{region 'Documentation'}
(*!
<summary>Immediately releases reservations for this Suite and all registered Test Cases.</summary>
<description>
Attempts every registered child and the own contribution even after an individual failure.
TRUE means all attempted releases succeeded; FALSE may mean partial release. Already released
contributions are not rolled back.

Does not change lifecycle states or stop cyclic child calls. During Reset-error finalization
it may free a child's budget before that child finishes; no new child requests may then be issued by
the completed Suite. This is failure cleanup, not normal admission.

Traverses the registered children only when finalized collection metadata is valid. Missing child interfaces or failed child releases make the result FALSE while remaining children and the own release are still attempted. The own zero contribution does not skip child traversal. This is not an initialization or resource-stop operation.
</description>
*)
{endregion}
// C0298: Reviewed compiler false positive in virtual/interface call-graph detection.
// Reported to Beckhoff; local suppression without a fabricated stack estimate.
{warning disable C0298}
METHOD PUBLIC FINAL FreeReservedEvents : BOOL //! TRUE when all subtree contributions were released; FALSE permits partial success.
VAR
    Index : LINT;
    Child : I_TestCase;
END_VAR
FreeReservedEvents := TRUE;
IF FCollectionConfiguration.IsValid THEN
    FOR Index := DINT_TO_LINT(FCollectionConfiguration.FirstIndex)
        TO DINT_TO_LINT(FCollectionConfiguration.FirstIndex) + UINT_TO_LINT(FCollectionConfiguration.Count) - 1 DO
        Child := GetTestCase(Index := LINT_TO_DINT(Index));
        IF Child = 0 THEN
            FreeReservedEvents := FALSE;
            CONTINUE;
        END_IF;
        IF NOT Child.FreeReservedEvents() THEN
            FreeReservedEvents := FALSE;
        END_IF;
    END_FOR;
END_IF;

IF UpdateEventReservation(EntryCount := 0,
    HeadroomEntryCount := 0,
    ChildEntryCount := 0) <> E_EventReservationResult.Accepted THEN
    FreeReservedEvents := FALSE;
END_IF;
{warning restore C0298}
END_METHOD

{region 'Documentation'}
(*!
<summary>Returns the common view from the typed owner collection without executing the
child.</summary>
*)
{endregion}
METHOD PUBLIC FINAL GetChild : I_Orchestratable //! Registered child interface at Index; zero for an invalid or unoccupied index.
VAR_INPUT
    Index : DINT; //! Original child-array index, not a registration ordinal; valid children occupy LowerBound through LowerBound + Count - 1.
END_VAR
GetChild := 0;
IF (ChildCount = 0) OR (Index < ChildArrayLowerBound)
    OR (DINT_TO_LINT(Index) >= DINT_TO_LINT(ChildArrayLowerBound) + UINT_TO_LINT(ChildCount)) THEN
    RETURN;
END_IF;
GetChild := GetTestCase(Index := Index);
END_METHOD

{region 'Documentation'}
(*!
<summary>Returns a registered child from the concrete owner's interface array.</summary>
<description>
Implement lookup in the same array configured by Configure, using its actual array index
rather than a hard-coded registration ordinal. Registration can reorder entries by slot.

Check the occupied range starting at ChildArrayLowerBound for ChildCount entries and return
zero outside it. Do not access unused capacity, execute the child, or cache a setup-time array
address. This abstract method has no base implementation.
</description>
*)
{endregion}
METHOD PUBLIC ABSTRACT GetTestCase : I_TestCase //! Registered child interface at Index; zero for an invalid or unoccupied index.
VAR_INPUT
    Index : DINT; //! Original child-array index, not a registration ordinal; valid children occupy LowerBound through LowerBound + Count - 1.
END_VAR
(* GetTestCase := 0;
IF (ChildCount = 0) OR (Index < ChildArrayLowerBound)
    OR (DINT_TO_LINT(Index) >= DINT_TO_LINT(ChildArrayLowerBound) + UINT_TO_LINT(ChildCount)) THEN
    RETURN;
END_IF;
GetTestCase := FTestCases[Index];
*)
END_METHOD

{region 'Documentation'}
(*!
<summary>Reports a detected Abort timeout until Initialize or entry into a new Reset.</summary>
<description>
An expired abort deadline finishes through Completing with Error. Escalation from Aborting to
AbortingFromError does not restart that deadline.
</description>
*)
{endregion}
{attribute 'monitoring' := 'call'}
PROPERTY PUBLIC HasAbortTimeout : BOOL //! Reports a detected Abort timeout until Initialize or entry into a new Reset.
GET // PUBLIC
HasAbortTimeout := FHasAbortTimeout;
END_GET
END_PROPERTY

{region 'Documentation'}
(*!
<summary>Reports the current owner error condition used by status projection.</summary>
*)
{endregion}
{attribute 'monitoring' := 'call'}
PROPERTY PUBLIC HasError : BOOL //! Reports the current owner error condition used by status projection.
GET // PUBLIC
HasError := FConfigError OR (FResult = E_Result.Error);
END_GET
END_PROPERTY

{region 'Documentation'}
(*!
<summary>Reports a detected Reset timeout until Initialize or entry into a new Reset.</summary>
<description>
The owner leaves a timed-out Reset through Completing to Completed with Error, not through
Abort. Capacity waiting or scenario cleanup remains part of the configured deadline.
</description>
*)
{endregion}
{attribute 'monitoring' := 'call'}
PROPERTY PUBLIC HasResetTimeout : BOOL //! Reports a detected Reset timeout until Initialize or entry into a new Reset.
GET // PUBLIC
HasResetTimeout := FHasResetTimeout;
END_GET
END_PROPERTY

{region 'Documentation'}
(*!
<summary>Reports a detected execution timeout until Initialize or entry into a new Reset.</summary>
<description>
The owner supervises its own execution deadline; the parent does not duplicate this check.
Invalid timer measurements report Framework errors without setting this timeout flag.
</description>
*)
{endregion}
{attribute 'monitoring' := 'call'}
PROPERTY PUBLIC HasTimeout : BOOL //! Reports a detected execution timeout until Initialize or entry into a new Reset.
GET // PUBLIC
HasTimeout := FHasTimeout;
END_GET
END_PROPERTY

{region 'Documentation'}
(*!
<summary>Establishes identity, invokes Configure, then validates the complete setup.</summary>
<description>
Called by the parent after Event Buffer startup initialization; clears only this owner's old
reservation. Configure rebuilds the child setup without releasing the previous registry. Parent is
not retained. Successful setup waits in Uninitialized for the parent's capacity-admitted Reset
request.

Reinitialization requires configuration reactivation or PLC Cold Reset followed by the
application's first-cycle initialization chain. Normal PLC Stop/Start and UnitTest Reset do not
rebuild configuration. Do not call Initialize as recovery during an active run.

The selected publisher must already be usable for configuration diagnostics. Failure leaves
IsInitialized FALSE; retained diagnostic identity is not proof of valid setup.
</description>
*)
{endregion}
METHOD PUBLIC FINAL Initialize : BOOL //! TRUE after successful identity and setup validation; FALSE leaves the object uninitialized.
VAR_INPUT
    Parent : I_RunControl; //! Owning Run Control with an established Name; read during Initialize, not retained.
    SuiteName : STRING(GVL_Constants.NameLength); //! Nonempty single name segment appended to Parent.Name; the complete name must fit NameLength.
    ResourceName : STRING(GVL_Constants.ResourceNameLength) := ''; //! Optional resource context for diagnostics; empty by default.
    Config : ST_TestSuiteConfig; //! Timeout configuration copied during initialization; all timeout values must be greater than zero.
END_VAR
VAR
    FullName : STRING(2 * GVL_Constants.NameLength + 1);
    EmptyStatus : ST_TestSuiteStatus;
    // SA0167: Setup-only builder; no state or binding survives this initialization call.
    {attribute 'analysis' := '-167'}
    Builder : TestSuiteConfigurationBuilder;
    EmptyCollectionConfiguration : ST_TestCaseCollectionConfig;
END_VAR
Initialize := FALSE;
FInitialized := FALSE;
FReservedEntryCount := 0;
FCollectionConfiguration := EmptyCollectionConfiguration;
FHasTimeout := FALSE;
FHasResetTimeout := FALSE;
FHasAbortTimeout := FALSE;
FState := E_State.Uninitialized;
FExecutionTimer.Reset();
FStateTimer.Start();
FAggregator.Reset();
FTestCaseCountInactive := 0;
FTestCaseCountIdle := 0;
FTestCaseCountRunning := 0;
FTestCaseCountCompleted := 0;
FTestCaseCountError := 0;
FCollectionValid := FALSE;
FChildrenError := FALSE;
FChildrenAborted := FALSE;
FChildrenCompleted := FALSE;
FChildrenAbortFinished := FALSE;
FCheckingInitialization := FALSE;
FConfigError := TRUE;
FName := SuiteName;
FResourceName := ResourceName;
FConfig := Config;
FResult := E_Result.NotEvaluated;
FStatus := EmptyStatus;
FStatus.Execution.Uninitialized := TRUE;
FStatus.Execution.ConfigError := TRUE;
FStatus.Execution.ExecutionStatus := E_ExecutionStatus.NotReady;
FMethodRequests.Start := FALSE;
FMethodRequests.Abort := FALSE;
FMethodRequests.Reset := FALSE;

IF Parent = 0 THEN
    PublishInitializationError(Message := 'Missing Run Control parent.');
    RETURN;
END_IF;
FullName := CONCAT(CONCAT(Parent.Name, '.'), SuiteName);
// SA0175: ASCII name contract; byte-based access is intentional and bounded.
{analysis -175}
FName := LEFT(FullName, UINT_TO_INT(GVL_Constants.NameLength));
{analysis +175}
IF NOT IsNameValid(Name := FullName, Depth := 2) THEN
    PublishInitializationError(Message := CONCAT('Invalid Test Suite name: ', FullName));
    RETURN;
END_IF;

Configure(Builder := Builder);
FCollectionConfiguration := Builder.Finalize();
IF NOT FCollectionConfiguration.IsValid THEN
    PublishInitializationError(Message := 'Invalid Test Case collection configuration.');
    RETURN;
END_IF;
IF FOrchestrator = 0 THEN
    FOrchestrator := FDefaultOrchestrator;
END_IF;

FCheckingInitialization := TRUE;
IF NOT FOrchestrator.Initialize(Collection := THIS^,
    Name := FName,
    ResourceName := FResourceName) THEN
    FCheckingInitialization := FALSE;
    PublishInitializationError(Message := 'Orchestrator initialization failed.');
    RETURN;
END_IF;

FConfigError := NOT CheckInitialization();
FCheckingInitialization := FALSE;
IF FConfigError THEN
    RETURN;
END_IF;

FInitialized := TRUE;
FStatus.Execution.ConfigError := FALSE;
FStatus.TestCaseCountTotal := ChildCount;
Initialize := TRUE;
END_METHOD

{region 'Documentation'}
(*!
<summary>Reports completed explicit abort, including the legacy Aborted state.</summary>
*)
{endregion}
{attribute 'monitoring' := 'call'}
PROPERTY PUBLIC IsAborted : BOOL //! Reports completed explicit abort, including the legacy Aborted state.
GET // PUBLIC
IsAborted := ((FState = E_State.Completed) AND (FResult = E_Result.Abort)) OR (FState = E_State.Aborted);
END_GET
END_PROPERTY

{region 'Documentation'}
(*!
<summary>Reports explicit or error-driven abort processing.</summary>
*)
{endregion}
{attribute 'monitoring' := 'call'}
PROPERTY PUBLIC IsAborting : BOOL //! Reports explicit or error-driven abort processing.
GET // PUBLIC
IsAborting := (FState = E_State.Aborting) OR (FState = E_State.AbortingFromError);
END_GET
END_PROPERTY

{region 'Documentation'}
(*!
<summary>Reports terminal completion independently of the result.</summary>
*)
{endregion}
{attribute 'monitoring' := 'call'}
PROPERTY PUBLIC IsComplete : BOOL //! Reports terminal completion independently of the result.
GET // PUBLIC
IsComplete := FState = E_State.Completed;
END_GET
END_PROPERTY

{region 'Documentation'}
(*!
<summary>Reports Idle state independently of readiness.</summary>
*)
{endregion}
{attribute 'monitoring' := 'call'}
PROPERTY PUBLIC IsIdle : BOOL //! Reports Idle state independently of readiness.
GET // PUBLIC
IsIdle := FState = E_State.Idle;
END_GET
END_PROPERTY

{region 'Documentation'}
(*!
<summary>Reports successful explicit identity, composition and configuration validation.</summary>
<description>
TRUE does not imply Idle or Ready. Successful Initialize still waits in Uninitialized for the
parent's capacity-admitted Reset.
</description>
*)
{endregion}
{attribute 'monitoring' := 'call'}
PROPERTY PUBLIC IsInitialized : BOOL //! Reports successful explicit identity, composition and configuration validation.
GET // PUBLIC
IsInitialized := FInitialized;
END_GET
END_PROPERTY

{region 'Documentation'}
(*!
<summary>Reports whether this owner can accept Start in Idle.</summary>
<description>
Requires successful initialization, valid configuration and collection, no owner Error, and
Orchestrator readiness with a neutral NotEvaluated helper result. The Orchestrator supplies the
child-readiness summary; IsInitialized or IsIdle alone is insufficient.
</description>
*)
{endregion}
{attribute 'monitoring' := 'call'}
PROPERTY PUBLIC IsReady : BOOL //! Reports whether this owner can accept Start in Idle.
GET // PUBLIC
IsReady := FALSE;
IF NOT FInitialized OR FConfigError OR (FResult = E_Result.Error) OR (FState <> E_State.Idle)
    OR NOT FCollectionValid THEN
    RETURN;
END_IF;
IsReady := FOrchestrator.IsReady
    AND (FOrchestrator.Result = E_Result.NotEvaluated);
END_GET
END_PROPERTY

{region 'Documentation'}
(*!
<summary>Reports active Reset processing.</summary>
*)
{endregion}
{attribute 'monitoring' := 'call'}
PROPERTY PUBLIC IsResetting : BOOL //! Reports active Reset processing.
GET // PUBLIC
IsResetting := FState = E_State.Reset;
END_GET
END_PROPERTY

{region 'Documentation'}
(*!
<summary>Checks a Suite transition without changing state or producing diagnostics.</summary>
*)
{endregion}
METHOD PRIVATE IsStateTransitionAllowed : BOOL //! TRUE when the requested state satisfies the current initialization, readiness, lifecycle and completion prerequisites.
VAR_INPUT
    NewState : E_State; //! Requested destination checked without changing state, result, timers or events.
END_VAR
IF NewState = E_State.Uninitialized THEN
    IsStateTransitionAllowed := TRUE;
    RETURN;
END_IF;
IF NOT FInitialized THEN
    IsStateTransitionAllowed := FALSE;
    RETURN;
END_IF;

CASE NewState OF
    E_State.Reset:
        IsStateTransitionAllowed := TRUE;
    E_State.Idle:
        IsStateTransitionAllowed := (FState = E_State.Reset) AND NOT FConfigError
            AND (FResult <> E_Result.Error) AND FCollectionValid
            AND FOrchestrator.IsResetFinished
            AND (FOrchestrator.Result = E_Result.NotEvaluated);
    E_State.Starting:
        IsStateTransitionAllowed := IsReady;
    E_State.Running:
        IsStateTransitionAllowed := (FState = E_State.Starting) AND (FResult <> E_Result.Error);
    E_State.Completing:
        CASE FState OF
            E_State.Uninitialized, E_State.Starting, E_State.Completed:
                IsStateTransitionAllowed := FALSE;
            E_State.Reset, E_State.Idle:
                IsStateTransitionAllowed := FResult = E_Result.Error;
            E_State.Running:
                IsStateTransitionAllowed := FChildrenCompleted AND (FResult <> E_Result.Error)
                    AND FOrchestrator.IsExecutionFinished;
            E_State.Aborting, E_State.AbortingFromError:
                IsStateTransitionAllowed := TRUE;
        ELSE
            IsStateTransitionAllowed := FResult = E_Result.Error;
        END_CASE;
    E_State.Completed:
        IsStateTransitionAllowed := FState = E_State.Completing;
    E_State.Aborting:
        IsStateTransitionAllowed := ((FState = E_State.Starting) OR (FState = E_State.Running))
            AND (FResult <> E_Result.Error);
    E_State.AbortingFromError:
        IsStateTransitionAllowed := ((FState = E_State.Starting) OR (FState = E_State.Running)
            OR (FState = E_State.Aborting)) AND (FResult = E_Result.Error);
ELSE
    IsStateTransitionAllowed := FALSE;
END_CASE;
END_METHOD

{region 'Documentation'}
(*!
<summary>Reports the active lifecycle, including finalization and abort processing.</summary>
*)
{endregion}
{attribute 'monitoring' := 'call'}
PROPERTY PUBLIC IsTestSuiteActive : BOOL //! Reports the active lifecycle, including finalization and abort processing.
GET // PUBLIC
IsTestSuiteActive := (FState = E_State.Starting) OR (FState = E_State.Running)
    OR (FState = E_State.Completing) OR IsAborting;
END_GET
END_PROPERTY

{region 'Documentation'}
(*!
<summary>Maps owner state and the current helper task; Reset finalization never selects Abort.</summary>
*)
{endregion}
METHOD PRIVATE MapOrchestratorTask : E_OrchestratorTask //! Helper task selected from State; Completing retains Execution/Abort, otherwise selects Idle.
VAR_INPUT
    State : E_State; //! Current owner lifecycle state after sequencing.
    CurrentTask : E_OrchestratorTask; //! Previously assigned helper task, retained during Completing only for Execution or Abort.
END_VAR
CASE State OF
    E_State.Reset:
        MapOrchestratorTask := E_OrchestratorTask.Reset;
    E_State.Starting, E_State.Running:
        MapOrchestratorTask := E_OrchestratorTask.Execution;
    E_State.Aborting, E_State.AbortingFromError:
        MapOrchestratorTask := E_OrchestratorTask.Abort;
    E_State.Completing:
        IF (CurrentTask = E_OrchestratorTask.Execution) OR (CurrentTask = E_OrchestratorTask.Abort) THEN
            MapOrchestratorTask := CurrentTask;
        ELSE
            MapOrchestratorTask := E_OrchestratorTask.Idle;
        END_IF;
ELSE
    MapOrchestratorTask := E_OrchestratorTask.Idle;
END_CASE;
END_METHOD

{region 'Documentation'}
(*!
<summary>Hierarchical identity retained for diagnostics, including rejected names.</summary>
*)
{endregion}
{attribute 'monitoring' := 'variable'}
PROPERTY PUBLIC Name : STRING(GVL_Constants.NameLength) //! Hierarchical identity retained for diagnostics, including rejected names.
GET // PUBLIC
Name := FName;
END_GET
END_PROPERTY

{region 'Documentation'}
(*!
<summary>Reads one child snapshot and accumulates lifecycle observations; invalid bindings invalidate the collection.</summary>
*)
{endregion}
METHOD PRIVATE ObserveTestCase : BOOL //! TRUE after reading an initialized child snapshot; FALSE clears ChildStatus and invalidates collection observations.
VAR_INPUT
    Child : I_TestCase; //! Borrowed Test Case interface; zero or uninitialized children invalidate collection observations.
END_VAR
VAR_OUTPUT
    ChildStatus : ST_TestCaseStatus; //! One child snapshot by value; empty on invalid binding. TRUE indicates binding validity rather than a successful verdict.
END_VAR
VAR
    ChildValid : BOOL;
    EmptyStatus : ST_TestCaseStatus;
END_VAR
ObserveTestCase := FALSE;
ChildValid := FALSE;
IF Child <> 0 THEN
    ChildValid := Child.IsInitialized;
END_IF;
IF NOT ChildValid THEN
    ChildStatus := EmptyStatus;
    FCollectionValid := FALSE;
    FChildrenCompleted := FALSE;
    FChildrenAbortFinished := FALSE;
    FChildrenError := TRUE;
    RETURN;
END_IF;

ChildStatus := Child.Status;
CASE ChildStatus.Execution.Result OF
    E_Result.NotEvaluated, E_Result.Passed, E_Result.Failed, E_Result.Abort, E_Result.Error:
        FChildrenError := FChildrenError OR (ChildStatus.Execution.Result = E_Result.Error);
ELSE
    FChildrenError := TRUE;
END_CASE;
FChildrenError := FChildrenError OR ChildStatus.Execution.Error OR ChildStatus.Execution.ConfigError
    OR (ChildStatus.Execution.ExecutionStatus = E_ExecutionStatus.Error);
FChildrenAborted := FChildrenAborted OR (ChildStatus.Execution.Result = E_Result.Abort);
FChildrenCompleted := FChildrenCompleted AND ChildStatus.Execution.Completed;
FChildrenAbortFinished := FChildrenAbortFinished
    AND (ChildStatus.Execution.Ready OR ChildStatus.Execution.Completed);
ObserveTestCase := TRUE;
END_METHOD

{region 'Documentation'}
(*!
<summary>Consumes same-task requests, reports each received request and prioritizes Reset &gt; Abort &gt; Start.</summary>
<description>
Discards requests before initialization; never changes lifecycle state.
</description>
*)
{endregion}
METHOD PRIVATE ProcessRequests
VAR_IN_OUT
    InputRequests : ST_Command; //! Same-task request mailbox consumed and cleared, including before successful initialization.
END_VAR
VAR_OUTPUT
    Requests : ST_Command; //! Qualified request snapshot with Reset over Abort over Start; all FALSE before initialization.
END_VAR
Requests.Reset := FALSE;
Requests.Abort := FALSE;
Requests.Start := FALSE;

IF NOT FInitialized THEN
    InputRequests.Reset := FALSE;
    InputRequests.Abort := FALSE;
    InputRequests.Start := FALSE;
    RETURN;
END_IF;

Requests.Reset := InputRequests.Reset;
Requests.Abort := InputRequests.Abort AND NOT InputRequests.Reset;
Requests.Start := InputRequests.Start AND NOT InputRequests.Abort AND NOT InputRequests.Reset;

IF InputRequests.Reset THEN
    PublishEvent(Event := CreateResetEvent(OwnerScope := E_OwnerScope.TestSuite,
        Name := FName,
        ResourceName := FResourceName,
        State := FState));
END_IF;

IF InputRequests.Abort THEN
    PublishEvent(Event := CreateAbortEvent(OwnerScope := E_OwnerScope.TestSuite,
        Name := FName,
        ResourceName := FResourceName,
        State := FState));
END_IF;

IF InputRequests.Start THEN
    PublishEvent(Event := CreateStartEvent(OwnerScope := E_OwnerScope.TestSuite,
        Name := FName,
        ResourceName := FResourceName,
        State := FState));
END_IF;

InputRequests.Reset := FALSE;
InputRequests.Abort := FALSE;
InputRequests.Start := FALSE;
END_METHOD

{region 'Documentation'}
(*!
<summary>Calls every owned Test Case exactly once per initialized cycle, including
Completed.</summary>
<description>
Do not gate child calls by parent state; child requests and lifecycle control their
work.
</description>
*)
{endregion}
METHOD PROTECTED ABSTRACT ProcessTestCases
(* Example: call every owned Test Case, including children not currently selected.
FTestCaseA();
FTestCaseB();
*)
END_METHOD

{region 'Documentation'}
(*!
<summary>Publishes through the selected instance publisher without owning buffer loss accounting.</summary>
*)
{endregion}
METHOD PRIVATE PublishEvent
VAR_INPUT
    Event : ST_Event; //! Payload forwarded once to the selected usable publisher, which assigns identity/time and accounts for loss.
END_VAR
EventPublisher.PublishEvent(Event := Event);
END_METHOD

{region 'Documentation'}
(*!
<summary>Emits a setup diagnostic without advancing lifecycle or changing the owner result.</summary>
*)
{endregion}
METHOD PRIVATE PublishInitializationError
VAR_INPUT
    Message : STRING(GVL_Constants.MessageLength); //! Setup diagnostic text sent through the required usable selected publisher without changing lifecycle or result.
END_VAR
EventPublisher.PublishEvent(Event := CreateFrameworkEvent(Name := FName,
    ResourceName := FResourceName,
    State := E_State.Uninitialized,
    Severity := E_EventSeverity.Error,
    Message := Message));
END_METHOD

{region 'Documentation'}
(*!
<summary>Records an Abort request for the next regular FB call.</summary>
<description>
Repeated positive calls coalesce in the same-task request storage. Processing consumes the
requests with priority Reset, Abort, Start; calls before successful initialization are discarded
when processed.

Abort requests controlled termination of execution, not Reset cancellation. The owner
lifecycle determines whether the request applies.
</description>
*)
{endregion}
METHOD PUBLIC RequestAbort
FMethodRequests.Abort := TRUE;
END_METHOD

{region 'Documentation'}
(*!
<summary>Records a Reset request for the next regular FB call.</summary>
<description>
Repeated positive calls coalesce in the same-task request storage. Processing consumes the
requests with priority Reset, Abort, Start; calls before successful initialization are discarded
when processed.

Lifecycle Reset preserves configuration and publisher binding. It is not reinitialization or
Event Buffer Reset; capacity admission belongs to the parent when this object is a child.

A new Reset entry returns from sequencing so the helper can initialize its Reset task before owner supervision reads its result. Further requests while Reset is active retain the deadline, held errors and dispatch progress and continue the regular clock, timeout and completion checks.
</description>
*)
{endregion}
METHOD PUBLIC RequestReset
FMethodRequests.Reset := TRUE;
END_METHOD

{region 'Documentation'}
(*!
<summary>Records a Start request for the next regular FB call.</summary>
<description>
Repeated positive calls coalesce in the same-task request storage. Processing consumes the
requests with priority Reset, Abort, Start; calls before successful initialization are discarded
when processed.

Start is accepted by the lifecycle only in ready Idle. Recording the request does not start
execution synchronously.
</description>
*)
{endregion}
METHOD PUBLIC RequestStart
FMethodRequests.Start := TRUE;
END_METHOD

{region 'Documentation'}
(*!
<summary>Own Suite reservation only; child contributions are not included.</summary>
*)
{endregion}
{attribute 'monitoring' := 'call'}
PROPERTY PUBLIC ReservedEntryCount : UINT //! Own Suite reservation only; child contributions are not included.
GET // PUBLIC
ReservedEntryCount := FReservedEntryCount;
END_GET
END_PROPERTY

{region 'Documentation'}
(*!
<summary>Adjusts this owner's reservation to its execution budget immediately.</summary>
<description>
Only this owner's contribution is reserved; child budgets are separate. Local contribution and
publisher accounting are updated together without a lifecycle transition.

Accepted permits dispatch; WaitingForCapacity is retryable under the owner's timeout; Error
denotes invalid setup or an impossible budget. Calling before initialization reports a Framework
error. Repeated success aligns the total rather than adding a second budget.
</description>
*)
{endregion}
METHOD PUBLIC FINAL ReserveExecutionEvents : E_EventReservationResult //! Accepted on success, WaitingForCapacity for retryable pressure, Error for invalid setup or an impossible budget.
ReserveExecutionEvents := E_EventReservationResult.Error;
IF NOT FInitialized THEN
    PublishEvent(Event := CreateFrameworkEvent(Name := FName,
        ResourceName := FResourceName,
        State := FState,
        Severity := E_EventSeverity.Error,
        Message := 'ReserveExecutionEvents requires an initialized Test Suite.'));
    RETURN;
END_IF;

ReserveExecutionEvents := UpdateEventReservation(EntryCount := GVL_Constants.TestSuiteExecutionEventCount,
    HeadroomEntryCount := Param_EventBuffer.EventBufferExecutionHeadroom,
    ChildEntryCount := 0);
END_METHOD

{region 'Documentation'}
(*!
<summary>Adjusts this owner's reservation for capacity-admitted Reset immediately.</summary>
<description>
Does not dispatch Reset or clear existing events. Shared headroom and one Test Case Reset
allowance participate in admission, not this owner's stored contribution.

Accepted, WaitingForCapacity and Error distinguish success, temporary pressure and invalid
setup. An uninitialized call reports a Framework error. Lifecycle Reset must not silently clear the
reservation.
</description>
*)
{endregion}
METHOD PUBLIC FINAL ReserveResetEvents : E_EventReservationResult //! Accepted on success, WaitingForCapacity for retryable pressure, Error for invalid setup or an impossible budget.
ReserveResetEvents := E_EventReservationResult.Error;
IF NOT FInitialized THEN
    PublishEvent(Event := CreateFrameworkEvent(Name := FName,
        ResourceName := FResourceName,
        State := FState,
        Severity := E_EventSeverity.Error,
        Message := 'ReserveResetEvents requires an initialized Test Suite.'));
    RETURN;
END_IF;

ReserveResetEvents := UpdateEventReservation(EntryCount := GVL_Constants.TestSuiteResetEventCount,
    HeadroomEntryCount := Param_EventBuffer.EventBufferResetHeadroom,
    ChildEntryCount := GVL_Constants.TestCaseResetEventCount);
END_METHOD

{region 'Documentation'}
(*!
<summary>Returns the owner result retained by the Suite lifecycle.</summary>
<description>
Ordinary execution remains NotEvaluated until finalization, while errors can be raised
earlier. Completed holds the final owner result even though child aggregation and status counters
continue refreshing. A new Reset clears the result.
</description>
*)
{endregion}
{attribute 'monitoring' := 'call'}
PROPERTY PUBLIC Result : E_Result //! Returns the owner result retained by the Suite lifecycle.
GET // PUBLIC
Result := FResult;
END_GET
END_PROPERTY

{region 'Documentation'}
(*!
<summary>Owns Suite transition decisions and timeout supervision; child request dispatch belongs to the shared Orchestrator.</summary>
<description>
A new Reset entry returns from sequencing so the helper can initialize its Reset task before owner supervision reads its result. Further requests while Reset is active retain the deadline, held errors and dispatch progress and continue the regular clock, timeout and completion checks.
</description>
*)
{endregion}
METHOD PRIVATE Sequencer
VAR_INPUT
    Requests : ST_Command; //! Consumed lifecycle request snapshot; only a new Reset entry returns before state-specific supervision.
END_VAR
IF NOT FInitialized THEN
    IF FState <> E_State.Uninitialized THEN
        ChangeState(NewState := E_State.Uninitialized);
    END_IF;
    RETURN;
END_IF;
IF Requests.Reset AND (FState <> E_State.Reset) THEN
    ChangeState(NewState := E_State.Reset);
    RETURN;
END_IF;

CASE FState OF
    E_State.Uninitialized:
        RETURN;

    E_State.Reset:
        IF NOT FCollectionValid THEN
            Error(Message := 'Registered Test Case collection is no longer valid.');
            ChangeState(NewState := E_State.Completing);
            RETURN;
        END_IF;
        IF NOT FStateTimer.IsValid THEN
            Error(Message := 'Task clock error during Test Suite reset.');
            ChangeState(NewState := E_State.Completing);
            RETURN;
        END_IF;
        IF FStateTimer.ElapsedLTime >= TIME_TO_LTIME(FConfig.ResetTimeout) THEN
            FHasResetTimeout := TRUE;
            PublishEvent(Event := CreateFrameworkEvent(Name := FName,
                ResourceName := FResourceName,
                State := FState,
                Severity := E_EventSeverity.Error,
                Message := 'Test Suite reset timeout reached.'));
            FResult := E_Result.Error;
            ChangeState(NewState := E_State.Completing);
            RETURN;
        END_IF;
        IF FOrchestrator.Result <> E_Result.NotEvaluated THEN
            Error(Message := 'Orchestrator failed during Test Suite reset.');
        END_IF;
        IF (FResult = E_Result.Error) AND FOrchestrator.IsResetFinished THEN
            ChangeState(NewState := E_State.Completing);
            RETURN;
        END_IF;
        IF FOrchestrator.IsResetFinished THEN
            ChangeState(NewState := E_State.Idle);
        END_IF;
        RETURN;

    E_State.Idle:
        IF NOT FCollectionValid THEN
            Error(Message := 'Registered Test Case collection is no longer valid.');
            ChangeState(NewState := E_State.Completing);
            RETURN;
        END_IF;
        IF FResult <> E_Result.Error THEN
            IF FChildrenError THEN
                Error(Message := 'A registered Test Case reported an error.');
            ELSIF FChildrenAborted AND (FResult <> E_Result.Abort) THEN
                Error(Message := 'Unexpected Test Case abort.');
            END_IF;
        END_IF;
        IF FResult = E_Result.Error THEN
            ChangeState(NewState := E_State.Completing);
            RETURN;
        END_IF;
        IF FOrchestrator.Result <> E_Result.NotEvaluated THEN
            Error(Message := 'Orchestrator is not ready for Test Suite start.');
            ChangeState(NewState := E_State.Completing);
            RETURN;
        END_IF;
        IF Requests.Start AND IsReady THEN
            ChangeState(NewState := E_State.Starting);
        END_IF;
        RETURN;

    E_State.Starting, E_State.Running:
        IF NOT FCollectionValid THEN
            Error(Message := 'Registered Test Case collection is no longer valid.');
            ChangeState(NewState := E_State.AbortingFromError);
            RETURN;
        END_IF;
        IF FResult <> E_Result.Error THEN
            IF FChildrenError THEN
                Error(Message := 'A registered Test Case reported an error.');
            ELSIF FChildrenAborted AND (FResult <> E_Result.Abort) THEN
                Error(Message := 'Unexpected Test Case abort.');
            END_IF;
        END_IF;
        IF FResult = E_Result.Error THEN
            ChangeState(NewState := E_State.AbortingFromError);
            RETURN;
        END_IF;
        IF FOrchestrator.Result = E_Result.Error THEN
            Error(Message := 'Orchestrator reported an execution error.');
            ChangeState(NewState := E_State.AbortingFromError);
            RETURN;
        END_IF;
        IF NOT FExecutionTimer.IsValid THEN
            Error(Message := 'Task clock error during Test Suite execution.');
            ChangeState(NewState := E_State.AbortingFromError);
            RETURN;
        END_IF;
        IF FExecutionTimer.ElapsedLTime >= TIME_TO_LTIME(FConfig.Timeout) THEN
            FHasTimeout := TRUE;
            Error(Message := 'Test Suite timeout reached.');
            ChangeState(NewState := E_State.AbortingFromError);
            RETURN;
        END_IF;
        IF Requests.Abort THEN
            ChangeState(NewState := E_State.Aborting);
            RETURN;
        END_IF;
        IF FState = E_State.Starting THEN
            ChangeState(NewState := E_State.Running);
            RETURN;
        END_IF;
        IF FChildrenCompleted AND FOrchestrator.IsExecutionFinished THEN
            ChangeState(NewState := E_State.Completing);
        END_IF;
        RETURN;

    E_State.Completing:
        ChangeState(NewState := E_State.Completed);
        RETURN;

    E_State.Completed:
        RETURN;

    E_State.Aborting, E_State.AbortingFromError:
        IF (FState = E_State.Aborting) AND NOT FCollectionValid THEN
            Error(Message := 'Registered Test Case collection is no longer valid.');
            ChangeState(NewState := E_State.AbortingFromError);
            RETURN;
        END_IF;
        IF FResult <> E_Result.Error THEN
            IF FChildrenError THEN
                Error(Message := 'A registered Test Case reported an error.');
            ELSIF FChildrenAborted AND (FResult <> E_Result.Abort) AND (FState <> E_State.Aborting) THEN
                Error(Message := 'Unexpected Test Case abort.');
            END_IF;
        END_IF;
        IF NOT FStateTimer.IsValid THEN
            PublishEvent(Event := CreateFrameworkEvent(Name := FName,
                ResourceName := FResourceName,
                State := FState,
                Severity := E_EventSeverity.Error,
                Message := 'Task clock error during Test Suite abort.'));
            FResult := E_Result.Error;
            ChangeState(NewState := E_State.Completing);
            RETURN;
        END_IF;
        IF FStateTimer.ElapsedLTime >= TIME_TO_LTIME(FConfig.AbortTimeout) THEN
            FHasAbortTimeout := TRUE;
            PublishEvent(Event := CreateFrameworkEvent(Name := FName,
                ResourceName := FResourceName,
                State := FState,
                Severity := E_EventSeverity.Error,
                Message := 'Test Suite abort timeout reached.'));
            FResult := E_Result.Error;
            ChangeState(NewState := E_State.Completing);
            RETURN;
        END_IF;
        IF (FState = E_State.Aborting) AND (FResult = E_Result.Error) THEN
            ChangeState(NewState := E_State.AbortingFromError);
            RETURN;
        END_IF;
        IF (FState = E_State.Aborting)
            AND (FOrchestrator.Result = E_Result.Error) THEN
            Error(Message := 'Orchestrator failed during Test Suite abort.');
            ChangeState(NewState := E_State.AbortingFromError);
            RETURN;
        END_IF;
        IF FChildrenAbortFinished AND FOrchestrator.IsAbortFinished THEN
            ChangeState(NewState := E_State.Completing);
        END_IF;
        RETURN;
ELSE
    IF NOT FCollectionValid THEN
        Error(Message := 'Registered Test Case collection is no longer valid.');
        ChangeState(NewState := E_State.Completing);
        RETURN;
    END_IF;
    IF FResult <> E_Result.Error THEN
        IF FChildrenError THEN
            Error(Message := 'A registered Test Case reported an error.');
        ELSIF FChildrenAborted AND (FResult <> E_Result.Abort) THEN
            Error(Message := 'Unexpected Test Case abort.');
        END_IF;
    END_IF;
    Error(Message := 'Unhandled Test Suite lifecycle state.');
    ChangeState(NewState := E_State.Completing);
END_CASE;
END_METHOD

{region 'Documentation'}
(*!
<summary>Current Suite lifecycle state.</summary>
*)
{endregion}
{attribute 'monitoring' := 'call'}
PROPERTY PUBLIC State : E_State //! Current Suite lifecycle state.
GET // PUBLIC
State := FState;
END_GET
END_PROPERTY

{region 'Documentation'}
(*!
<summary>Returns the latest cyclic owner-status snapshot.</summary>
<description>
Status is refreshed on every FB call, including Uninitialized and Completed. Runtime uses
TIME; child counters may continue changing after final event publication. Reading this property
performs no child processing and does not republish final events.
</description>
*)
{endregion}
PROPERTY PUBLIC Status : ST_TestSuiteStatus //! Returns the latest cyclic owner-status snapshot.
GET // PUBLIC
Status := FStatus;
END_GET
END_PROPERTY

{region 'Documentation'}
(*!
<summary>Checks own budget plus unreserved child allowance before changing either count.</summary>
<description>
Zero releases without capacity gating.

A zero target with no held contribution succeeds without publisher access. A nonzero held contribution is released through FreeReservedSpace without free-capacity gating. Positive targets check actual publisher validity/accounting and permanent capacity for target plus child allowance plus headroom. Temporary free capacity uses aggregate minus old own contribution plus target plus child allowance plus headroom. Even unchanged or reduced positive targets must pass this check. Only the Suite contribution changes; child allowance remains shared unreserved capacity. Failure leaves both ledgers unchanged.
</description>
*)
{endregion}
METHOD PRIVATE UpdateEventReservation : E_EventReservationResult //! Accepted after aligning the own contribution, WaitingForCapacity for temporary pressure, Error for invalid prerequisites or an impossible budget.
VAR_INPUT
    EntryCount : UINT; //! Target total own reservation, not an additional delta; zero releases the entire own contribution.
    HeadroomEntryCount : UINT; //! Shared unreserved producer headroom used in permanent and temporary capacity checks for positive targets.
    ChildEntryCount : UINT; //! Unreserved child allowance used in both permanent and temporary capacity checks; never added to the Suite's own ledger.
END_VAR
VAR
    Publisher : I_EventPublisher;
    RequiredCapacity : UDINT;
    RequiredFreeEntries : UDINT;
END_VAR
UpdateEventReservation := E_EventReservationResult.Error;
IF (EntryCount = 0) AND (FReservedEntryCount = 0) THEN
    UpdateEventReservation := E_EventReservationResult.Accepted;
    RETURN;
END_IF;

Publisher := EventPublisher;

IF EntryCount = 0 THEN
    IF Publisher.FreeReservedSpace(EntryCount := FReservedEntryCount,
        OwnerReservedEntryCount := FReservedEntryCount) THEN
        UpdateEventReservation := E_EventReservationResult.Accepted;
    END_IF;
    RETURN;
END_IF;

IF NOT Publisher.IsValid THEN
    RETURN;
END_IF;
RequiredCapacity := UINT_TO_UDINT(EntryCount)
    + UINT_TO_UDINT(ChildEntryCount)
    + UINT_TO_UDINT(HeadroomEntryCount);
IF RequiredCapacity > UINT_TO_UDINT(Publisher.Capacity) THEN
    RETURN;
END_IF;
IF FReservedEntryCount > Publisher.ReservedEntryCount THEN
    RETURN;
END_IF;

RequiredFreeEntries := UINT_TO_UDINT(Publisher.ReservedEntryCount)
    - UINT_TO_UDINT(FReservedEntryCount)
    + UINT_TO_UDINT(EntryCount)
    + UINT_TO_UDINT(ChildEntryCount)
    + UINT_TO_UDINT(HeadroomEntryCount);
IF RequiredFreeEntries > UINT_TO_UDINT(Publisher.FreeEntryCount) THEN
    UpdateEventReservation := E_EventReservationResult.WaitingForCapacity;
    RETURN;
END_IF;

IF EntryCount < FReservedEntryCount THEN
    IF Publisher.FreeReservedSpace(EntryCount := FReservedEntryCount - EntryCount,
        OwnerReservedEntryCount := FReservedEntryCount) THEN
        UpdateEventReservation := E_EventReservationResult.Accepted;
    END_IF;
    RETURN;
END_IF;

IF Publisher.ReserveSpace(EntryCount := EntryCount - FReservedEntryCount,
    HeadroomEntryCount := HeadroomEntryCount,
    OwnerReservedEntryCount := FReservedEntryCount) THEN
    UpdateEventReservation := E_EventReservationResult.Accepted;
ELSE
    UpdateEventReservation := E_EventReservationResult.WaitingForCapacity;
END_IF;
END_METHOD

{region 'Documentation'}
(*!
<summary>Applies owner result semantics to the current child aggregate without changing lifecycle state.</summary>
*)
{endregion}
METHOD PRIVATE UpdateResult
VAR
    OrchestratorResult : E_Result;
END_VAR
IF FState = E_State.Uninitialized THEN
    FResult := E_Result.NotEvaluated;
    RETURN;
END_IF;
IF (FState = E_State.Reset) OR (FState = E_State.Completed) OR (FResult = E_Result.Error) THEN
    RETURN;
END_IF;

IF NOT FCollectionValid THEN
    Error(Message := 'Registered Test Case collection is no longer valid.');
    RETURN;
END_IF;
IF FChildrenError OR (FAggregator.Result = E_Result.Error) THEN
    Error(Message := 'A registered Test Case reported an error.');
    RETURN;
END_IF;
OrchestratorResult := FOrchestrator.Result;
IF OrchestratorResult = E_Result.Error THEN
    Error(Message := 'Orchestrator reported an error.');
    RETURN;
END_IF;
IF (FAggregator.Result = E_Result.Abort)
    AND (FResult <> E_Result.Abort) AND (FState <> E_State.Aborting) THEN
    Error(Message := 'Unexpected Test Case abort.');
    RETURN;
END_IF;

CASE FState OF
    E_State.Idle, E_State.Starting, E_State.Running:
        FResult := E_Result.NotEvaluated;
    E_State.Aborting:
        FResult := E_Result.Abort;
    E_State.AbortingFromError:
        FResult := E_Result.Error;
    E_State.Completing:
        IF FResult = E_Result.Abort THEN
            RETURN;
        END_IF;
        IF (FResult = E_Result.Failed) OR (FAggregator.Result = E_Result.Failed) THEN
            FResult := E_Result.Failed;
            RETURN;
        END_IF;
        FResult := E_Result.Passed;
ELSE
    Error(Message := 'Unhandled Test Suite lifecycle state.');
END_CASE;
END_METHOD

{region 'Documentation'}
(*!
<summary>Projects lifecycle, runtime and internally collected counters on every FB call, including Completed.</summary>
*)
{endregion}
METHOD PRIVATE UpdateStatus
VAR
    Execution : ST_ExecutionStatus;
END_VAR
Execution.State := FState;
Execution.Result := FResult;
Execution.ConfigError := FConfigError;
CASE FState OF
    E_State.Uninitialized:
        Execution.ExecutionStatus := E_ExecutionStatus.NotReady;
        Execution.Uninitialized := TRUE;
    E_State.Reset:
        Execution.ExecutionStatus := E_ExecutionStatus.Reset;
    E_State.Idle:
        Execution.ExecutionStatus := E_ExecutionStatus.Idle;
        Execution.Ready := IsReady;
    E_State.Starting:
        Execution.ExecutionStatus := E_ExecutionStatus.Starting;
    E_State.Running:
        Execution.ExecutionStatus := E_ExecutionStatus.Running;
        Execution.Running := TRUE;
    E_State.Completing:
        Execution.ExecutionStatus := E_ExecutionStatus.Completing;
    E_State.Completed:
        Execution.ExecutionStatus := E_ExecutionStatus.Completed;
        Execution.Completed := TRUE;
        Execution.Aborted := FResult = E_Result.Abort;
    E_State.Aborting, E_State.AbortingFromError:
        Execution.ExecutionStatus := E_ExecutionStatus.Aborting;
ELSE
    Execution.ExecutionStatus := E_ExecutionStatus.Error;
END_CASE;
Execution.Error := HasError;
FStatus.Execution := Execution;
FStatus.Runtime := FExecutionTimer.ElapsedTime;
FStatus.TestCaseCountTotal := ChildCount;
FStatus.TestCaseCountInactive := FTestCaseCountInactive;
FStatus.TestCaseCountIdle := FTestCaseCountIdle;
FStatus.TestCaseCountRunning := FTestCaseCountRunning;
FStatus.TestCaseCountCompleted := FTestCaseCountCompleted;
FStatus.TestCaseCountError := FTestCaseCountError;
FStatus.TestCaseCountPassed := FAggregator.PassedCount;
FStatus.TestCaseCountFailed := FAggregator.FailedCount;
END_METHOD

END_FUNCTION_BLOCK

// ---- Framework/TestSuites/POU/TestSuiteConfigurationBuilder.TcPOU
{region 'Documentation'}
(*!
<summary>Setup-only configuration: Initialize through Finalize requires stable array/child storage.</summary>
<description>
No FB body call is required. Finalize discards the temporary array pointer on either outcome.
At most 65535 children can be registered; Initialize clears the array after validating mode and capacity.


The returned configuration describes the owner's actual array; Finalize does not copy child storage or make it immutable. Keep that array, child instances and assigned slots stable for the complete execution lifetime. Do not retain a temporary builder passed to Configure. Setup clears array capacity and scans/shifts registered entries; it is configuration work, not cyclic scheduling.
</description>
*)
{endregion}
FUNCTION_BLOCK TestSuiteConfigurationBuilder
VAR
    FInitialized : BOOL;
    FEntries : POINTER TO I_TestCase;
    FFinalized : BOOL;
    FRegistrationError : BOOL;
    FConfiguration : ST_TestCaseCollectionConfig;
END_VAR

VAR CONSTANT
    MaxCount : UINT := 65535;
END_VAR

{region 'Documentation'}
(*!
<summary>Number of registered entries, contiguous from FirstIndex.</summary>
*)
{endregion}
{attribute 'monitoring' := 'call'}
PROPERTY PUBLIC Count : UINT //! Number of registered entries, contiguous from FirstIndex.
GET // PUBLIC
Count := FConfiguration.Count;
END_GET
END_PROPERTY

{region 'Documentation'}
(*!
<summary>Finalizes validation and releases the array binding; repeated calls return the same configuration.</summary>
<description>
Rejects empty collections, latched errors and invalid slots. Serial slots follow registration order, Parallel uses slot one, and ParallelSlots must form consecutive positive groups beginning at one. The temporary array pointer is discarded on success and failure; repeated calls return the frozen configuration. Child initialization is checked later by the Suite, not here.
</description>
*)
{endregion}
METHOD PUBLIC Finalize : ST_TestCaseCollectionConfig //! Finalized bounds, count and mode; IsValid determines whether the configuration can be used.
VAR
    Offset : DINT;
    PreviousSlot : UDINT;
    Slot : UDINT;
    Child : I_TestCase;
END_VAR
IF FFinalized THEN
    Finalize := FConfiguration;
    RETURN;
END_IF;

IF NOT FInitialized OR FRegistrationError OR (FEntries = 0) OR (FConfiguration.Count = 0) THEN
    FConfiguration.IsValid := FALSE;
    FEntries := 0;
    FFinalized := TRUE;
    Finalize := FConfiguration;
    RETURN;
END_IF;

PreviousSlot := 0;
FOR Offset := 0 TO UINT_TO_DINT(FConfiguration.Count) - 1 DO
    Child := FEntries[Offset];
    IF Child = 0 THEN
        FRegistrationError := TRUE;
        EXIT;
    END_IF;
    Slot := UINT_TO_UDINT(Child.ExecutionSlot);
    IF (Slot = 0) OR (Slot < PreviousSlot) OR (Slot > PreviousSlot + 1)
        OR ((FConfiguration.Mode = E_OrchestrationMode.Serial) AND (Slot <> DINT_TO_UDINT(Offset) + 1))
        OR ((FConfiguration.Mode = E_OrchestrationMode.Parallel) AND (Slot <> 1)) THEN
        FRegistrationError := TRUE;
        EXIT;
    END_IF;
    PreviousSlot := Slot;
END_FOR;

FConfiguration.IsValid := NOT FRegistrationError;
FEntries := 0;
FFinalized := TRUE;
Finalize := FConfiguration;
END_METHOD

{region 'Documentation'}
(*!
<summary>Actual lower bound of the supplied array.</summary>
*)
{endregion}
{attribute 'monitoring' := 'call'}
PROPERTY PUBLIC FirstIndex : DINT //! Actual lower bound of the supplied array.
GET // PUBLIC
FirstIndex := FConfiguration.FirstIndex;
END_GET
END_PROPERTY

{region 'Documentation'}
(*!
<summary>Starts a new build and clears the supplied array; bounds and mode remain fixed until Finalize.</summary>
<description>
Validate mode and positive physical capacity before clearing entries; rejected prerequisites leave the array untouched. Occupied entries form a contiguous prefix at the actual lower bound. Initialize starts a fresh build after prior success or failure; at most 65535 children can be registered even in a larger array.
</description>
*)
{endregion}
METHOD PUBLIC Initialize
VAR_INPUT
    Mode : E_OrchestrationMode; //! Scheduling strategy fixed for this build; Register is for Serial/Parallel, RegisterWithSlot for ParallelSlots.
END_VAR
VAR_IN_OUT
    TestCases : ARRAY[*] OF I_TestCase; //! Owner-held array cleared and filled by the builder; storage must stay fixed through Finalize and registered children must outlive execution.
END_VAR
VAR
    Index : LINT;
    Capacity : LINT;
END_VAR
FInitialized := FALSE;
FEntries := 0;
FFinalized := FALSE;
FRegistrationError := FALSE;
FConfiguration.IsValid := FALSE;
FConfiguration.Count := 0;
FConfiguration.FirstIndex := LOWER_BOUND(TestCases, 1);
FConfiguration.LastIndex := UPPER_BOUND(TestCases, 1);
FConfiguration.Mode := Mode;

IF (Mode <> E_OrchestrationMode.Serial)
    AND (Mode <> E_OrchestrationMode.Parallel)
    AND (Mode <> E_OrchestrationMode.ParallelSlots) THEN
    FRegistrationError := TRUE;
    RETURN;
END_IF;

Capacity := DINT_TO_LINT(FConfiguration.LastIndex) - DINT_TO_LINT(FConfiguration.FirstIndex) + 1;
IF Capacity <= 0 THEN
    FRegistrationError := TRUE;
    RETURN;
END_IF;

FOR Index := DINT_TO_LINT(FConfiguration.FirstIndex) TO DINT_TO_LINT(FConfiguration.LastIndex) DO
    TestCases[LINT_TO_DINT(Index)] := 0;
END_FOR;
FEntries := ADR(TestCases[FConfiguration.FirstIndex]);
FInitialized := TRUE;
END_METHOD

{region 'Documentation'}
(*!
<summary>Validates before mutation, inserts the child and sets its effective slot.</summary>
*)
{endregion}
METHOD PRIVATE Insert : BOOL //! TRUE after insertion and slot assignment; FALSE latches a registration error without adding an entry.
VAR_INPUT
    TestCase : I_TestCase; //! Unique nonzero Test Case interface whose instance must outlive the finalized collection.
    ExecutionSlot : UINT; //! Positive effective slot; stable insertion preserves registration order within equal slots.
END_VAR
VAR
    Offset : DINT;
    InsertOffset : DINT;
    Child : I_TestCase;
END_VAR
Insert := FALSE;
IF NOT FInitialized OR FRegistrationError OR (FEntries = 0) OR (TestCase = 0) OR (ExecutionSlot = 0) THEN
    FRegistrationError := TRUE;
    RETURN;
END_IF;
IF (FConfiguration.Count = MaxCount)
    OR (UINT_TO_LINT(FConfiguration.Count) >= DINT_TO_LINT(FConfiguration.LastIndex) - DINT_TO_LINT(FConfiguration.FirstIndex) + 1) THEN
    FRegistrationError := TRUE;
    RETURN;
END_IF;

InsertOffset := UINT_TO_DINT(FConfiguration.Count);
FOR Offset := 0 TO UINT_TO_DINT(FConfiguration.Count) - 1 DO
    Child := FEntries[Offset];
    IF (Child = 0) OR (Child = TestCase) THEN
        FRegistrationError := TRUE;
        RETURN;
    END_IF;
    IF (InsertOffset = UINT_TO_DINT(FConfiguration.Count)) AND (Child.ExecutionSlot > ExecutionSlot) THEN
        InsertOffset := Offset;
    END_IF;
END_FOR;
IF FEntries[FConfiguration.Count] <> 0 THEN
    FRegistrationError := TRUE;
    RETURN;
END_IF;

TestCase.ExecutionSlot := ExecutionSlot;
FOR Offset := UINT_TO_DINT(FConfiguration.Count) TO InsertOffset + 1 BY -1 DO
    FEntries[Offset] := FEntries[Offset - 1];
END_FOR;
FEntries[InsertOffset] := TestCase;
FConfiguration.Count := FConfiguration.Count + 1;
Insert := TRUE;
END_METHOD

{region 'Documentation'}
(*!
<summary>Finalize has completed, independently of validation success.</summary>
*)
{endregion}
{attribute 'monitoring' := 'call'}
PROPERTY PUBLIC IsFinalized : BOOL //! Finalize has completed, independently of validation success.
GET // PUBLIC
IsFinalized := FFinalized;
END_GET
END_PROPERTY

{region 'Documentation'}
(*!
<summary>Finalization succeeded; FALSE before Finalize.</summary>
*)
{endregion}
{attribute 'monitoring' := 'call'}
PROPERTY PUBLIC IsValid : BOOL //! Finalization succeeded; FALSE before Finalize.
GET // PUBLIC
IsValid := FConfiguration.IsValid;
END_GET
END_PROPERTY

{region 'Documentation'}
(*!
<summary>Actual upper bound, including unused capacity.</summary>
*)
{endregion}
{attribute 'monitoring' := 'call'}
PROPERTY PUBLIC LastIndex : DINT //! Actual upper bound, including unused capacity.
GET // PUBLIC
LastIndex := FConfiguration.LastIndex;
END_GET
END_PROPERTY

{region 'Documentation'}
(*!
<summary>Mode selected by Initialize.</summary>
*)
{endregion}
{attribute 'monitoring' := 'call'}
PROPERTY PUBLIC Mode : E_OrchestrationMode //! Mode selected by Initialize.
GET // PUBLIC
Mode := FConfiguration.Mode;
END_GET
END_PROPERTY

{region 'Documentation'}
(*!
<summary>Appends a unique child in Serial or Parallel mode and assigns its effective slot.</summary>
<description>
Serial assigns increasing slots; Parallel uses slot one. A rejection before finalization latches a build error until another Initialize. After Finalize this method returns FALSE without altering the frozen configuration or latching a new error.
</description>
*)
{endregion}
METHOD PUBLIC Register : BOOL //! TRUE when the child was registered; FALSE adds no entry; pre-finalization rejection latches a build error.
VAR_INPUT
    TestCase : I_TestCase; //! Nonzero child interface to register once; its instance must outlive the registered collection.
END_VAR
VAR
    Slot : UINT;
END_VAR
Register := FALSE;
IF FFinalized THEN
    RETURN;
END_IF;
IF (FConfiguration.Mode <> E_OrchestrationMode.Serial)
    AND (FConfiguration.Mode <> E_OrchestrationMode.Parallel) THEN
    FRegistrationError := TRUE;
    RETURN;
END_IF;

Slot := 1;
IF FConfiguration.Mode = E_OrchestrationMode.Serial THEN
    IF FConfiguration.Count = MaxCount THEN
        FRegistrationError := TRUE;
        RETURN;
    END_IF;
    Slot := FConfiguration.Count + 1;
END_IF;
Register := Insert(TestCase := TestCase,
    ExecutionSlot := Slot);
END_METHOD

{region 'Documentation'}
(*!
<summary>Registers a unique child in ParallelSlots mode, stably inserting by positive slot.</summary>
<description>
Only for ParallelSlots. Positive slots are stably sorted into the array; Finalize checks consecutive groups beginning at one. Rejection before finalization latches a build error; after Finalize FALSE does not change the frozen outcome.
</description>
*)
{endregion}
METHOD PUBLIC RegisterWithSlot : BOOL //! TRUE when the child was registered; FALSE adds no entry; pre-finalization rejection latches a build error.
VAR_INPUT
    TestCase : I_TestCase; //! Nonzero child interface to register once; its instance must outlive the registered collection.
    ExecutionSlot : UINT; //! Positive slot number for ParallelSlots registration; children sharing a slot may overlap, with at most one new Start admitted per helper call.
END_VAR
RegisterWithSlot := FALSE;
IF FFinalized THEN
    RETURN;
END_IF;
IF FConfiguration.Mode <> E_OrchestrationMode.ParallelSlots THEN
    FRegistrationError := TRUE;
    RETURN;
END_IF;
RegisterWithSlot := Insert(TestCase := TestCase,
    ExecutionSlot := ExecutionSlot);
END_METHOD

END_FUNCTION_BLOCK

// ---- Framework/EventBuffer/POU/AggregationEvents/CreateTestSuiteAggregationEvent.TcPOU
{region 'Documentation'}
(*!
<summary>Constructs a Test Suite aggregation event from an already aggregated status snapshot.</summary>
<description>
Runtime is rendered as unsigned milliseconds; the caller owns publication.


Compact JSON fields are total, inactive, idle, running, completed, passed, failed, error and runtime. Counts and runtime are unsigned decimal numbers. This formats the supplied snapshot without validating completion or recomputing aggregation; the owner controls finalization order and publication.
</description>
*)
{endregion}
FUNCTION CreateTestSuiteAggregationEvent : ST_Event //! Constructed event value; not published. The publisher assigns SequenceId and Timestamp.
VAR_INPUT
    Name : STRING(GVL_Constants.NameLength); //! Hierarchical owner name used to identify events; must satisfy the naming contract.
    ResourceName : STRING(GVL_Constants.ResourceNameLength) := ''; //! Optional resource context for diagnostics; empty by default.
    Status : ST_TestSuiteStatus; //! Already aggregated owner status snapshot; the function formats it without observing children.
END_VAR
VAR
    RuntimeMilliseconds : UDINT;
END_VAR

RuntimeMilliseconds := TIME_TO_UDINT(Status.Runtime);

CreateTestSuiteAggregationEvent.SequenceId := 0;
CreateTestSuiteAggregationEvent.Timestamp := 0;
CreateTestSuiteAggregationEvent.OwnerScope := E_OwnerScope.TestSuite;
CreateTestSuiteAggregationEvent.EventType := E_EventType.Aggregation;
CreateTestSuiteAggregationEvent.Severity := SelectResultSeverity(Result := Status.Execution.Result);
CreateTestSuiteAggregationEvent.Name := Name;
CreateTestSuiteAggregationEvent.ResourceName := ResourceName;
CreateTestSuiteAggregationEvent.State := Status.Execution.State;
CreateTestSuiteAggregationEvent.Result := Status.Execution.Result;

CreateTestSuiteAggregationEvent.Message := CONCAT(STR1 := '{"total":',
    STR2 := UINT_TO_STRING(Status.TestCaseCountTotal));
CreateTestSuiteAggregationEvent.Message := CONCAT(STR1 := CreateTestSuiteAggregationEvent.Message,
    STR2 := ',"inactive":');
CreateTestSuiteAggregationEvent.Message := CONCAT(STR1 := CreateTestSuiteAggregationEvent.Message,
    STR2 := UINT_TO_STRING(Status.TestCaseCountInactive));
CreateTestSuiteAggregationEvent.Message := CONCAT(STR1 := CreateTestSuiteAggregationEvent.Message,
    STR2 := ',"idle":');
CreateTestSuiteAggregationEvent.Message := CONCAT(STR1 := CreateTestSuiteAggregationEvent.Message,
    STR2 := UINT_TO_STRING(Status.TestCaseCountIdle));
CreateTestSuiteAggregationEvent.Message := CONCAT(STR1 := CreateTestSuiteAggregationEvent.Message,
    STR2 := ',"running":');
CreateTestSuiteAggregationEvent.Message := CONCAT(STR1 := CreateTestSuiteAggregationEvent.Message,
    STR2 := UINT_TO_STRING(Status.TestCaseCountRunning));
CreateTestSuiteAggregationEvent.Message := CONCAT(STR1 := CreateTestSuiteAggregationEvent.Message,
    STR2 := ',"completed":');
CreateTestSuiteAggregationEvent.Message := CONCAT(STR1 := CreateTestSuiteAggregationEvent.Message,
    STR2 := UINT_TO_STRING(Status.TestCaseCountCompleted));
CreateTestSuiteAggregationEvent.Message := CONCAT(STR1 := CreateTestSuiteAggregationEvent.Message,
    STR2 := ',"passed":');
CreateTestSuiteAggregationEvent.Message := CONCAT(STR1 := CreateTestSuiteAggregationEvent.Message,
    STR2 := UINT_TO_STRING(Status.TestCaseCountPassed));
CreateTestSuiteAggregationEvent.Message := CONCAT(STR1 := CreateTestSuiteAggregationEvent.Message,
    STR2 := ',"failed":');
CreateTestSuiteAggregationEvent.Message := CONCAT(STR1 := CreateTestSuiteAggregationEvent.Message,
    STR2 := UINT_TO_STRING(Status.TestCaseCountFailed));
CreateTestSuiteAggregationEvent.Message := CONCAT(STR1 := CreateTestSuiteAggregationEvent.Message,
    STR2 := ',"error":');
CreateTestSuiteAggregationEvent.Message := CONCAT(STR1 := CreateTestSuiteAggregationEvent.Message,
    STR2 := UINT_TO_STRING(Status.TestCaseCountError));
CreateTestSuiteAggregationEvent.Message := CONCAT(STR1 := CreateTestSuiteAggregationEvent.Message,
    STR2 := ',"runtime":');
CreateTestSuiteAggregationEvent.Message := CONCAT(STR1 := CreateTestSuiteAggregationEvent.Message,
    STR2 := UDINT_TO_STRING(RuntimeMilliseconds));
CreateTestSuiteAggregationEvent.Message := CONCAT(STR1 := CreateTestSuiteAggregationEvent.Message, STR2 := '}');

END_FUNCTION

// ---- SelfTests/TestCases/TestSuite_Smoke/Test_Smoke.TcPOU
{region 'Documentation'}
(*!
<summary>Exercises the successful framework lifecycle with one Boolean Assertion.</summary>
*)
{endregion}
FUNCTION_BLOCK Test_Smoke EXTENDS TestCaseBase
VAR
    FSuccess : AssertTrue;
    FActual : BOOL;
    FCheckPerformed : BOOL;
END_VAR

SUPER^();

{region 'Documentation'}
(*!
<summary>Contributes the one Assertion without executing or resetting it.</summary>
*)
{endregion}
METHOD PROTECTED AggregateResults
VAR_INPUT
    Aggregator : I_ResultAggregator; //! Borrowed result sink owned by the outer Test Case; add this test's checking Assertions without resetting or retaining the sink.
END_VAR
Aggregator.AddProvider(Provider := FSuccess);
END_METHOD

{region 'Documentation'}
(*!
<summary>Includes the owned Assertion in the base initialization checks.</summary>
*)
{endregion}
METHOD PROTECTED CheckInitialization : BOOL //! TRUE when the inherited initialization check and this concrete fixture check both accept the setup.
CheckInitialization := FALSE;
IF NOT SUPER^.CheckInitialization() THEN
    RETURN;
END_IF;
IF NOT FSuccess.IsInitialized THEN
    RETURN;
END_IF;

CheckInitialization := TRUE;
END_METHOD

{region 'Documentation'}
(*!
<summary>Initializes the smoke scenario and its single Assertion.</summary>
*)
{endregion}
METHOD PROTECTED Configure
FPreparationStateCount := 0;
FTestStateCount := 1;
FActual := FALSE;
FCheckPerformed := FALSE;

FSuccess.Initialize(Parent := THIS^,
    AssertionName := 'Success');
END_METHOD

{region 'Documentation'}
(*!
<summary>Completes enabled aborts; the smoke scenario owns no resource actions.</summary>
*)
{endregion}
METHOD PROTECTED ProcessAbort
VAR_INPUT
    Enable : BOOL; //! Phase permission supplied by the owning Test Case; FALSE does not authorize progression, while observation may continue.
END_VAR
IF Enable THEN
    CompleteAbort();
END_IF;
END_METHOD

{region 'Documentation'}
(*!
<summary>Calls the Assertion even while disabled and records an actual evaluation.</summary>
*)
{endregion}
METHOD PROTECTED ProcessAssertions
VAR_INPUT
    Enable : BOOL; //! Phase permission supplied by the owning Test Case; FALSE does not authorize progression, while observation may continue.
END_VAR
FSuccess(Enable := Enable,
    State := State,
    IN := FActual);

IF Enable AND FSuccess.EvaluationActive THEN
    FCheckPerformed := TRUE;
END_IF;
END_METHOD

{region 'Documentation'}
(*!
<summary>No Preparation stage is configured for this smoke scenario.</summary>
*)
{endregion}
METHOD PROTECTED ProcessPreparations
VAR_INPUT
    // SA0033: Required override signature; this scenario has no preparation work.
    {attribute 'analysis' := '-33'}
    Enable : BOOL; //! Phase permission supplied by the owning Test Case; FALSE does not authorize progression, while observation may continue.
END_VAR
END_METHOD

{region 'Documentation'}
(*!
<summary>Clears scenario progress and requests Assertion reset before returning to Idle.</summary>
*)
{endregion}
METHOD PROTECTED ProcessReset
FActual := FALSE;
FCheckPerformed := FALSE;
FSuccess.Reset();
CompleteReset();
END_METHOD

{region 'Documentation'}
(*!
<summary>Supplies the success value, then completes on the call after evaluation.</summary>
*)
{endregion}
METHOD PROTECTED ProcessTests
VAR_INPUT
    Enable : BOOL; //! Phase permission supplied by the owning Test Case; FALSE does not authorize progression, while observation may continue.
END_VAR
IF NOT Enable THEN
    RETURN;
END_IF;

IF FCheckPerformed THEN
    CompleteTests();
ELSE
    FActual := TRUE;
END_IF;
END_METHOD

END_FUNCTION_BLOCK

// ---- Framework/TestCases/POU/TestCaseBase.TcPOU
{region 'Documentation'}
(*!
<summary>Base-owned Test Case lifecycle with scenario-specific Preparation, test and Assertion
hooks.</summary>
<description>
The Suite calls Initialize before regular processing. Implement Configure, ProcessReset,
ProcessAbort, ProcessPreparations, ProcessTests, ProcessAssertions and AggregateResults; the
concrete FB body calls SUPER^() once per task cycle.

The base owns requests, transitions, timers, result interpretation and lifecycle events.
Completed skips processing hooks, but existing Assertion results and status counters are still
collected. Do not implement a second owner lifecycle in the concrete body.
</description>
*)
{endregion}
FUNCTION_BLOCK ABSTRACT TestCaseBase IMPLEMENTS I_TestCase
VAR CONSTANT
    StateCountNotConfigured : INT := -1;
END_VAR
VAR
    /// Instance binding; derived test adapters may assign it before first use.
    FEventPublisher : I_EventPublisher;
    FName : STRING(GVL_Constants.NameLength);
    FResourceName : STRING(GVL_Constants.ResourceNameLength);
    FConfig : ST_TestCaseConfig;
    FInitialized : BOOL;
FHasTimeout : BOOL;
FHasPreparationTimeout : BOOL;
FHasResetTimeout : BOOL;
FHasAbortTimeout : BOOL;
    FConfigError : BOOL;
    FExecutionSlot : UINT;
    FReservedEntryCount : UINT;
    FState : E_State := E_State.Uninitialized;
    FResult : E_Result := E_Result.NotEvaluated;
    FStatus : ST_TestCaseStatus;
    FPreparationStatus : ST_PreparationStatus;
    FPreparationStateCount : INT := StateCountNotConfigured;
    FTestStateCount : INT := StateCountNotConfigured;
    FExecutionTimer : Stopwatch;
    FStateTimer : Stopwatch;
    FMethodRequests: ST_Command;
    FAggregator : ResultAggregator;
END_VAR
VAR_TEMP
    Requests : ST_Command;
END_VAR

ProcessRequests(InputRequests := FMethodRequests, Requests => Requests);

FExecutionTimer.Update();
FStateTimer.Update();

Sequencer(Requests := Requests);

IF IsInitialized THEN
    IF IsResetting THEN
        FPreparationStatus.State := E_State.Uninitialized;
        FPreparationStatus.ExecutionStatus := E_ExecutionStatus.Unknown;
        FPreparationStatus.Ready := FALSE;
        FPreparationStatus.Running := FALSE;
        FPreparationStatus.Completed := FALSE;
        FPreparationStatus.Error := FALSE;
        UpdateStatus();
        ProcessReset();
    END_IF;

    IF FState <> E_State.Completed THEN
        ProcessAbort(Enable := IsAborting);

        ProcessPreparations(Enable := IsPreparationActive);
        ProcessTests(Enable := IsTestingActive);
        ProcessAssertions(Enable := IsTestingActive);
    END_IF;

    FAggregator.Reset();
    AggregateResults(Aggregator := FAggregator);
END_IF;

UpdateResult();
UpdateStatus();
EmitFinalizationEvents();

{region 'Documentation'}
(*!
<summary>Contributes every owned Assertion result exactly once to the current collection.</summary>
<description>
Called on every initialized FB call, including Completed and inactive phases. AddProvider or
AddResult contributes one counted Assertion; include inactive Assertions too.

The base resets the aggregator before the call and subsequently derives owner result, status
counters and finalization events. Do not reset or retain the passed interface, execute Assertions,
publish findings or latch another result here. This abstract hook has no base implementation.
</description>
*)
{endregion}
METHOD PROTECTED ABSTRACT AggregateResults
VAR_INPUT
    Aggregator : I_ResultAggregator; //! Owner-held contribution interface; add each child once without resetting or retaining this interface.
END_VAR
(* Example: add each owned Assertion once; do not reset the aggregator.
Aggregator.AddProvider(Provider := MyAssertion);
Aggregator.AddProvider(Provider := MyOtherAssertion);
*)
END_METHOD

{region 'Documentation'}
(*!
<summary>Applies permitted transitions; rejection holds state/timers and reports a diagnostic or Error according to the current lifecycle phase.</summary>
*)
{endregion}
METHOD PRIVATE ChangeState
VAR_INPUT
    NewState : E_State; //! Requested lifecycle destination; identical state is a no-op and rejection leaves state and timers unchanged.
END_VAR
IF NewState = FState THEN
    RETURN;
END_IF;

IF NOT IsStateTransitionAllowed(NewState := NewState) THEN
    CASE FState OF
        E_State.Uninitialized:
            RETURN;

        E_State.Completed:
            PublishEvent(Event := CreateInvalidStateTransitionEvent(OwnerScope := E_OwnerScope.TestCase,
                Name := FName,
                ResourceName := FResourceName,
                StateOld := FState,
                StateNew := NewState));
    ELSE
        IF FResult <> E_Result.Error THEN
            PublishEvent(Event := CreateInvalidStateTransitionEvent(OwnerScope := E_OwnerScope.TestCase,
                Name := FName,
                ResourceName := FResourceName,
                StateOld := FState,
                StateNew := NewState));
        END_IF;
        FResult := E_Result.Error;
    END_CASE;
    RETURN;
END_IF;

CASE NewState OF
    E_State.Uninitialized:
        FInitialized := FALSE;
        FResult := E_Result.NotEvaluated;
        FAggregator.Reset();
        FExecutionTimer.Reset();
        FStateTimer.Reset();

    E_State.Reset:
        FHasTimeout := FALSE;
        FHasPreparationTimeout := FALSE;
        FHasResetTimeout := FALSE;
        FHasAbortTimeout := FALSE;
        IF IsTestCaseActive THEN
            PublishEvent(Event := CreateResetWarningEvent(OwnerScope := E_OwnerScope.TestCase,
                Name := FName,
                ResourceName := FResourceName,
                State := FState));
        END_IF;
        FResult := E_Result.NotEvaluated;
        FAggregator.Reset();
        FExecutionTimer.Reset();
        FStateTimer.Start();

    E_State.Idle:
        FStateTimer.Reset();

    E_State.Starting:
        FExecutionTimer.Start();
        FStateTimer.Reset();

    E_State.Preparing..(E_State.Running - 1),
    E_State.Running..(E_State.Completing - 1):
        FStateTimer.Start();

    E_State.Aborting:
        FResult := E_Result.Abort;
        FExecutionTimer.Stop();
        FStateTimer.Start();

    E_State.AbortingFromError:
        FResult := E_Result.Error;
        FExecutionTimer.Stop();
        IF FState <> E_State.Aborting THEN
            FStateTimer.Start();
        END_IF;

    E_State.Completing:
        FExecutionTimer.Stop();
        FStateTimer.Reset();

    E_State.Completed:
        FStateTimer.Reset();
ELSE
    RETURN;
END_CASE;

PublishEvent(Event := CreateStateTransitionEvent(OwnerScope := E_OwnerScope.TestCase,
    Name := FName,
    ResourceName := FResourceName,
    StateOld := FState,
    StateNew := NewState));
FState := NewState;
END_METHOD

{region 'Documentation'}
(*!
<summary>Validates configured state counts and positive timeouts after Configure.</summary>
<description>
An override must call SUPER^.CheckInitialization(), retain failure, and additionally validate
its owned setup, including Assertion initialization. Return FALSE for any invalid prerequisite; do
not turn a failed base check into success.

The base reports its first failed check as a Framework diagnostic. Initialization remains
unsuccessful when validation fails.
</description>
*)
{endregion}
METHOD PROTECTED CheckInitialization : BOOL //! TRUE when the configured setup is valid; FALSE reports invalid setup and prevents initialization.
CheckInitialization := FALSE;

IF FPreparationStateCount = StateCountNotConfigured THEN
    PublishEvent(Event := CreateFrameworkEvent(Name := FName,
        ResourceName := FResourceName,
        State := FState,
        Severity := E_EventSeverity.Error,
        Message := 'Preparation state count was not configured.'));
    RETURN;
END_IF;

IF FTestStateCount = StateCountNotConfigured THEN
    PublishEvent(Event := CreateFrameworkEvent(Name := FName,
        ResourceName := FResourceName,
        State := FState,
        Severity := E_EventSeverity.Error,
        Message := 'Test state count was not configured.'));
    RETURN;
END_IF;

IF (FPreparationStateCount < 0)
    OR (FPreparationStateCount > E_State.Running - E_State.Preparing) THEN
    PublishEvent(Event := CreateFrameworkEvent(Name := FName,
        ResourceName := FResourceName,
        State := FState,
        Severity := E_EventSeverity.Error,
        Message := CONCAT('Invalid Preparation state count = ', INT_TO_STRING(FPreparationStateCount))));
    RETURN;
END_IF;

IF (FTestStateCount < 1)
    OR (FTestStateCount > E_State.Completing - E_State.Running) THEN
    PublishEvent(Event := CreateFrameworkEvent(Name := FName,
        ResourceName := FResourceName,
        State := FState,
        Severity := E_EventSeverity.Error,
        Message := CONCAT('Invalid Test state count = ', INT_TO_STRING(FTestStateCount))));
    RETURN;
END_IF;

IF (FConfig.Timeout = T#0MS) OR (FConfig.PreparationTimeout = T#0MS)
    OR (FConfig.ResetTimeout = T#0MS) OR (FConfig.AbortTimeout = T#0MS) THEN
    PublishEvent(Event := CreateFrameworkEvent(Name := FName,
        ResourceName := FResourceName,
        State := FState,
        Severity := E_EventSeverity.Error,
        Message := 'Timeout, PreparationTimeout, ResetTimeout and AbortTimeout must be greater than zero.'));
    RETURN;
END_IF;

CheckInitialization := TRUE;
END_METHOD

{region 'Documentation'}
(*!
<summary>Acknowledges finished cleanup and enters Completing immediately.</summary>
<description>
Call only during IsAborting, including the error-driven abort phase. The existing Abort or
Error result is preserved by finalization. The base enforces AbortTimeout even if the implementation
never acknowledges completion.
</description>
*)
{endregion}
METHOD PROTECTED CompleteAbort
IF NOT (IsAborting) THEN
    Error(Message := 'CompleteAbort called outside its lifecycle phase.');
    RETURN;
END_IF;
ChangeState(NewState := E_State.Completing);
END_METHOD

{region 'Documentation'}
(*!
<summary>Ends the active Preparation phase immediately by entering Running.</summary>
<description>
The concrete scenario must establish that its target is reached before calling. Held owner,
aggregate or Preparation Error prevents normal completion. The transition requires the
stored Completed flag as well as an error-free Preparation snapshot.

Following hooks observe the changed phase immediately. Alternatively, the Sequencer advances
from Starting or Preparing when the supplied Preparation snapshot already reports Completed.
</description>
*)
{endregion}
METHOD PROTECTED CompletePreparations
IF NOT IsPreparationActive THEN
    Error(Message := 'CompletePreparations called outside its lifecycle phase.');
    RETURN;
END_IF;
IF (FResult = E_Result.Error) OR (FAggregator.Result = E_Result.Error) THEN
    Error(Message := 'Test Case evaluation reported Error.');
    RETURN;
END_IF;

IF FPreparationStatus.Error THEN
    Error(Message := 'Preparation reported Error.');
    RETURN;
END_IF;
ChangeState(NewState := E_State.Running);
END_METHOD

{region 'Documentation'}
(*!
<summary>Acknowledges completed reset work.</summary>
<description>
Call only in Reset. Without a held Error, the owner enters Idle; with Error, it enters
Completing and then Completed, never an abort phase. Readiness in Idle still depends on the
effective IsReady implementation.

ResetTimeout bounds missing acknowledgement. This operation does not reinitialize
configuration or release event reservations.
</description>
*)
{endregion}
METHOD PROTECTED CompleteReset
IF NOT (FState = E_State.Reset) THEN
    Error(Message := 'CompleteReset called outside its lifecycle phase.');
    RETURN;
END_IF;
IF FResult = E_Result.Error THEN
    ChangeState(NewState := E_State.Completing);
    RETURN;
END_IF;
ChangeState(NewState := E_State.Idle);
END_METHOD

{region 'Documentation'}
(*!
<summary>Ends the active Test phase immediately by entering Completing.</summary>
<description>
Call only after scenario completion and error checks. Held owner or aggregate Error prevents
normal completion. Subsequent hooks in the same FB call see the new state; in particular
ProcessAssertions receives the updated IsTestingActive value.

This method does not evaluate Assertions or publish final results itself. The base collects
results and emits finalization events later in the call.
</description>
*)
{endregion}
METHOD PROTECTED CompleteTests
IF NOT IsTestingActive THEN
    Error(Message := 'CompleteTests called outside its lifecycle phase.');
    RETURN;
END_IF;
IF (FResult = E_Result.Error) OR (FAggregator.Result = E_Result.Error) THEN
    Error(Message := 'Test Case evaluation reported Error.');
    RETURN;
END_IF;

ChangeState(NewState := E_State.Completing);
END_METHOD

{region 'Documentation'}
(*!
<summary>Configures this concrete scenario and initializes its owned components.</summary>
<description>
Called synchronously after identity validation on every Initialize. Set both
FPreparationStateCount and FTestStateCount explicitly: zero Preparations is valid; at least one Test
state is required.

Counts describe the longest finite lifecycle path and must fit the corresponding E_State
intervals. Initialize Assertions with Parent := THIS^ and unique local names; preserve child
initialization failures for CheckInitialization.

This abstract hook has no base implementation to call. Do not perform cyclic test work
here.

Clear application-owned transient progress and pending resource commands here. Disabled hooks
may run after successful Initialize while the owner still waits for its parent's Reset; they must
already be passive.
</description>
*)
{endregion}
METHOD PROTECTED ABSTRACT Configure
(* Set counts for the longest finite path of this concrete scenario.
FPreparationStateCount := 0;
FTestStateCount := 1;
MyAssertion.Initialize(Parent := THIS^, AssertionName := 'MyAssertion');
Check MyAssertion.IsInitialized in CheckInitialization.
Initialize any owned components and retain their initialization failures for CheckInitialization.
*)
END_METHOD

{region 'Documentation'}
(*!
<summary>Publishes Result and Aggregation while in Completing, after result and status updates.</summary>
<description>
The base's single-call Completing phase supplies one-shot publication without a separate latch: the following regular sequencing call enters Completed. Result and Aggregation use the final status from this call. Failed insertion is accounted for by the publisher, with no retry here.
</description>
*)
{endregion}
METHOD PRIVATE EmitFinalizationEvents
IF (FState <> E_State.Completing) THEN
    RETURN;
END_IF;

PublishEvent(Event := CreateResultEvent(OwnerScope := E_OwnerScope.TestCase,
    Name := FName,
    ResourceName := FResourceName,
    State := FState,
    Result := FResult,
    Message := ''));
PublishEvent(Event := CreateTestCaseAggregationEvent(Name := FName, ResourceName := FResourceName, Status := FStatus));
END_METHOD

{region 'Documentation'}
(*!
<summary>Ignores Uninitialized and Completed; reports only before Result becomes Error.</summary>
<description>
Latches Error without leaving Reset or Idle; active execution enters controlled error
termination.
</description>
*)
{endregion}
METHOD PROTECTED Error
VAR_INPUT
    Message : STRING(GVL_Constants.MessageLength); //! Diagnostic text copied into the event within MessageLength.
END_VAR
IF (FState = E_State.Uninitialized) OR (FState = E_State.Completed) THEN
    RETURN;
END_IF;

IF FResult <> E_Result.Error THEN
    PublishEvent(Event := CreateFrameworkEvent(Name := FName,
        ResourceName := FResourceName,
        State := FState,
        Severity := E_EventSeverity.Error,
        Message := Message));
END_IF;

FResult := E_Result.Error;
IF (FState = E_State.Reset) OR (FState = E_State.Idle) THEN
    RETURN;
END_IF;
ChangeState(NewState := E_State.AbortingFromError);
END_METHOD

{region 'Documentation'}
(*!
<summary>Returns this instance's retained event-publication service.</summary>
<description>
If the local binding is zero, the getter takes GVL_EventBuffer.Publisher on access. An
established binding is retained; Initialize and lifecycle Reset do not replace it.

The default must be bound before first diagnostic use. Controlled test adapters may assign the
protected field before use. This getter performs no event publication, lifecycle processing or
reservation change.
</description>
*)
{endregion}
{attribute 'monitoring' := 'variable'}
PROPERTY PUBLIC EventPublisher : I_EventPublisher //! Returns this instance's retained event-publication service.
GET // PUBLIC
IF FEventPublisher = 0 THEN
    FEventPublisher := GVL_EventBuffer.Publisher;
END_IF;
EventPublisher := FEventPublisher;
END_GET
END_PROPERTY

{region 'Documentation'}
(*!
<summary>Suite-assigned slot; set only during configuration. Initialize and Reset retain
it.</summary>
*)
{endregion}
{attribute 'monitoring' := 'call'}
PROPERTY PUBLIC ExecutionSlot : UINT //! Suite-assigned slot; set only during configuration. Initialize and Reset retain it.
GET // PUBLIC
ExecutionSlot := FExecutionSlot;
END_GET
SET // PUBLIC
FExecutionSlot := ExecutionSlot;
END_SET
END_PROPERTY

{region 'Documentation'}
(*!
<summary>Releases the entire own reservation; zero is already successful, even before
initialization.</summary>
*)
{endregion}
METHOD PUBLIC FINAL FreeReservedEvents : BOOL //! TRUE when the own reservation is released or already zero; FALSE retains the unresolved contribution.
FreeReservedEvents := UpdateEventReservation(EntryCount := 0,
    HeadroomEntryCount := 0,
    ConcurrentEntryCount := 0) = E_EventReservationResult.Accepted;
END_METHOD

{region 'Documentation'}
(*!
<summary>Reports a detected Abort timeout until Initialize or entry into a new Reset.</summary>
<description>
An expired abort deadline finishes through Completing with Error. Escalation from Aborting to
AbortingFromError does not restart that deadline.
</description>
*)
{endregion}
{attribute 'monitoring' := 'call'}
PROPERTY PUBLIC HasAbortTimeout : BOOL //! Reports a detected Abort timeout until Initialize or entry into a new Reset.
GET // PUBLIC
HasAbortTimeout := FHasAbortTimeout;
END_GET
END_PROPERTY

{region 'Documentation'}
(*!
<summary>Reports the current owner error condition used by status projection.</summary>
*)
{endregion}
{attribute 'monitoring' := 'call'}
PROPERTY PUBLIC HasError : BOOL //! Reports the current owner error condition used by status projection.
GET // PUBLIC
HasError := FConfigError OR (FResult = E_Result.Error);
CASE FState OF
    E_State.Uninitialized, E_State.Reset, E_State.Idle, E_State.Starting,
    E_State.Completing, E_State.Completed, E_State.Aborting, E_State.AbortingFromError:
        RETURN;
ELSE
    HasError := HasError OR NOT (IsPreparationActive OR IsTestingActive);
END_CASE;
END_GET
END_PROPERTY

{region 'Documentation'}
(*!
<summary>Reports a detected Preparation timeout until Initialize or entry into a new
Reset.</summary>
*)
{endregion}
{attribute 'monitoring' := 'call'}
PROPERTY PUBLIC HasPreparationTimeout : BOOL //! Reports a detected Preparation timeout until Initialize or entry into a new Reset.
GET // PUBLIC
HasPreparationTimeout := FHasPreparationTimeout;
END_GET
END_PROPERTY

{region 'Documentation'}
(*!
<summary>Reports a detected Reset timeout until Initialize or entry into a new Reset.</summary>
<description>
The owner leaves a timed-out Reset through Completing to Completed with Error, not through
Abort. The deadline starts on entry into Reset and bounds scenario cleanup; the parent supervises earlier reservation waiting.
</description>
*)
{endregion}
{attribute 'monitoring' := 'call'}
PROPERTY PUBLIC HasResetTimeout : BOOL //! Reports a detected Reset timeout until Initialize or entry into a new Reset.
GET // PUBLIC
HasResetTimeout := FHasResetTimeout;
END_GET
END_PROPERTY

{region 'Documentation'}
(*!
<summary>Reports a detected execution timeout until Initialize or entry into a new Reset.</summary>
<description>
The owner supervises its own execution deadline; the parent does not duplicate this check.
Invalid timer measurements report Framework errors without setting this timeout flag.
</description>
*)
{endregion}
{attribute 'monitoring' := 'call'}
PROPERTY PUBLIC HasTimeout : BOOL //! Reports a detected execution timeout until Initialize or entry into a new Reset.
GET // PUBLIC
HasTimeout := FHasTimeout;
END_GET
END_PROPERTY

{region 'Documentation'}
(*!
<summary>Reinitializes the owner; validates identity before child setup and configuration
afterwards.</summary>
<description>
Clears its own old reservation after Event Buffer startup initialization; no old contribution
is released. Called by the parent at PLC start. Parent is not retained; the Suite-assigned
ExecutionSlot is retained. Successful setup waits in Uninitialized for the parent's
capacity-admitted Reset request.

Reinitialization requires configuration reactivation or PLC Cold Reset followed by the
application's first-cycle initialization chain. Normal PLC Stop/Start and UnitTest Reset do not
rebuild configuration. Do not call Initialize as recovery during an active run.

The selected publisher must already be usable for configuration diagnostics. Failure leaves
IsInitialized FALSE; retained diagnostic identity is not proof of valid setup.
</description>
*)
{endregion}
// C0298: Reviewed compiler false positive in virtual/interface call-graph detection.
// Reported to Beckhoff; local suppression without a fabricated stack estimate.
{warning disable C0298}
METHOD PUBLIC FINAL Initialize : BOOL //! TRUE after successful identity and setup validation; FALSE leaves the object uninitialized.
VAR_INPUT
    Parent : I_TestSuite; //! Owning Test Suite with an established Name; read during Initialize, not retained.
    TestName : STRING(GVL_Constants.NameLength); //! Nonempty single name segment appended to Parent.Name; the complete name must fit NameLength.
    ResourceName : STRING(GVL_Constants.ResourceNameLength) := ''; //! Optional resource context for diagnostics; empty by default.
    Config : ST_TestCaseConfig; //! Timeout configuration copied during initialization; all timeout values must be greater than zero.
END_VAR
VAR
    ParentName : STRING(GVL_Constants.NameLength);
    FullName : STRING(2 * GVL_Constants.NameLength + 1);
END_VAR
Initialize := FALSE;
FHasTimeout := FALSE;
FHasPreparationTimeout := FALSE;
FHasResetTimeout := FALSE;
FHasAbortTimeout := FALSE;
FInitialized := FALSE;
FReservedEntryCount := 0;
FConfigError := TRUE;
FState := E_State.Uninitialized;
FResult := E_Result.NotEvaluated;
FPreparationStateCount := StateCountNotConfigured;
FTestStateCount := StateCountNotConfigured;
FMethodRequests.Start := FALSE;
FMethodRequests.Abort := FALSE;
FMethodRequests.Reset := FALSE;
FAggregator.Reset();
FExecutionTimer.Reset();
FStateTimer.Reset();
FPreparationStatus.State := E_State.Uninitialized;
FPreparationStatus.ExecutionStatus := E_ExecutionStatus.Unknown;
FPreparationStatus.Ready := FALSE;
FPreparationStatus.Running := FALSE;
FPreparationStatus.Completed := FALSE;
FPreparationStatus.Error := FALSE;

IF Parent = 0 THEN
    FName := '';
    FResourceName := '';
    PublishEvent(Event := CreateFrameworkEvent(Name := TestName,
        ResourceName := ResourceName,
        State := FState,
        Severity := E_EventSeverity.Error,
        Message := 'Missing Test Suite parent.'));
    UpdateStatus();
    RETURN;
END_IF;

ParentName := Parent.Name;
FullName := CONCAT(CONCAT(ParentName, '.'), TestName);
// SA0175: ASCII name contract; byte-based access is intentional and bounded.
{analysis -175}
FName := LEFT(FullName, UINT_TO_INT(GVL_Constants.NameLength));
{analysis +175}
FResourceName := ResourceName;
FConfig := Config;

IF NOT IsNameValid(Name := FullName, Depth := 3) THEN
    PublishEvent(Event := CreateFrameworkEvent(Name := FName,
        ResourceName := FResourceName,
        State := FState,
        Severity := E_EventSeverity.Error,
        Message := CONCAT('Invalid Test Case name: ', FullName)));
    UpdateStatus();
    RETURN;
END_IF;

Configure();
FConfigError := NOT CheckInitialization();
FInitialized := NOT FConfigError;
Initialize := FInitialized;
UpdateStatus();
{warning restore C0298}
END_METHOD

{region 'Documentation'}
(*!
<summary>Reports a completed Abort result or the legacy Aborted state.</summary>
*)
{endregion}
{attribute 'monitoring' := 'call'}
PROPERTY PUBLIC IsAborted : BOOL //! Reports a completed Abort result or the legacy Aborted state.
GET // PUBLIC
IsAborted := ((FState = E_State.Completed) And (FResult = E_Result.Abort)) OR (FState = E_State.Aborted);
END_GET
END_PROPERTY

{region 'Documentation'}
(*!
<summary>Reports an active abort phase, including abort handling caused by Error.</summary>
*)
{endregion}
{attribute 'monitoring' := 'call'}
PROPERTY PUBLIC IsAborting : BOOL //! Reports an active abort phase, including abort handling caused by Error.
GET // PUBLIC
IsAborting := (FState = E_State.Aborting) OR (FState = E_State.AbortingFromError);
END_GET
END_PROPERTY

{region 'Documentation'}
(*!
<summary>Reports that the lifecycle has reached Completed, independent of its result.</summary>
*)
{endregion}
{attribute 'monitoring' := 'call'}
PROPERTY PUBLIC IsComplete : BOOL //! Reports that the lifecycle has reached Completed, independent of its result.
GET // PUBLIC
IsComplete := (FState = E_State.Completed);
END_GET
END_PROPERTY

{region 'Documentation'}
(*!
<summary>Reports Idle state independently of readiness.</summary>
*)
{endregion}
{attribute 'monitoring' := 'call'}
PROPERTY PUBLIC IsIdle : BOOL //! Reports Idle state independently of readiness.
GET // PUBLIC
IsIdle := FState = E_State.Idle;
END_GET
END_PROPERTY

{region 'Documentation'}
(*!
<summary>Reports successful explicit initialization.</summary>
*)
{endregion}
{attribute 'monitoring' := 'call'}
PROPERTY PUBLIC IsInitialized : BOOL //! Reports successful explicit initialization.
GET // PUBLIC
IsInitialized := FInitialized;
END_GET
END_PROPERTY

{region 'Documentation'}
(*!
<summary>Reports membership in the configured Preparation-state interval.</summary>
*)
{endregion}
{attribute 'monitoring' := 'call'}
PROPERTY PUBLIC IsPreparationActive : BOOL //! Reports membership in the configured Preparation-state interval.
GET // PUBLIC
IsPreparationActive := (FState >= E_State.Preparing) AND (FState < E_State.Preparing + FPreparationStateCount);
END_GET
END_PROPERTY

{region 'Documentation'}
(*!
<summary>Reports the effective Test Case start permission.</summary>
<description>
The base requires initialized, valid setup, Idle and no held Error. Override only when
additional resource or scenario prerequisites exist and combine them with SUPER^.IsReady. The status
snapshot uses this same effective property.
</description>
*)
{endregion}
{attribute 'monitoring' := 'call'}
PROPERTY PUBLIC IsReady : BOOL //! Reports the effective Test Case start permission.
GET // PUBLIC
IsReady := FInitialized AND NOT FConfigError AND (FState = E_State.Idle)
    AND (FResult <> E_Result.Error);
END_GET
END_PROPERTY

{region 'Documentation'}
(*!
<summary>Reports an active Reset phase.</summary>
*)
{endregion}
{attribute 'monitoring' := 'call'}
PROPERTY PUBLIC IsResetting : BOOL //! Reports an active Reset phase.
GET // PUBLIC
IsResetting := (FState = E_State.Reset);
END_GET
END_PROPERTY

{region 'Documentation'}
(*!
<summary>Checks the requested transition without changing state, result, timers or events.</summary>
*)
{endregion}
METHOD PRIVATE IsStateTransitionAllowed : BOOL //! TRUE when NewState satisfies the current lifecycle, configured state ranges and completion/error prerequisites.
VAR_INPUT
    NewState : E_State; //! Requested destination checked without changing state, result, timers or events.
END_VAR
IsStateTransitionAllowed := TRUE;
IF NewState = FState THEN
    RETURN;
END_IF;

CASE NewState OF
    E_State.Uninitialized:
        IsStateTransitionAllowed := TRUE;

    E_State.Reset:
        IsStateTransitionAllowed := FInitialized;

    E_State.Idle:
        IsStateTransitionAllowed := (FState = E_State.Reset) AND FInitialized AND NOT FConfigError;

    E_State.Starting:
        IsStateTransitionAllowed := (FState = E_State.Idle) AND IsReady;

    E_State.Preparing..(E_State.Running - 1):
        IsStateTransitionAllowed := FInitialized AND
            (NewState < E_State.Preparing + FPreparationStateCount) AND
            (((FState = E_State.Starting) AND (NewState = E_State.Preparing)) OR
            (IsPreparationActive AND (NewState = FState + 1)));
        IF FPreparationStatus.Error THEN
            IsStateTransitionAllowed := FALSE;
        END_IF;

    E_State.Running..(E_State.Completing - 1):
        IF NewState = E_State.Running THEN
            IsStateTransitionAllowed := FInitialized AND (FTestStateCount > 0) AND
                (((FState = E_State.Starting) AND (FPreparationStateCount = 0)) OR
                (((FState = E_State.Starting) OR IsPreparationActive) AND
                FPreparationStatus.Completed AND NOT FPreparationStatus.Error));
        ELSE
            IsStateTransitionAllowed := FInitialized AND IsTestingActive AND
                (NewState = FState + 1) AND
                (NewState < E_State.Running + FTestStateCount);
        END_IF;

    E_State.Completing:
        IsStateTransitionAllowed := IsTestingActive OR IsAborting
            OR ((FState = E_State.Reset) AND (FResult = E_Result.Error));

    E_State.Completed:
        IsStateTransitionAllowed := FState = E_State.Completing;

    E_State.Aborting:
        IsStateTransitionAllowed := ((FState = E_State.Starting) OR IsPreparationActive OR IsTestingActive)
            AND (FResult <> E_Result.Error) AND (FAggregator.Result <> E_Result.Error);

    E_State.AbortingFromError:
        IsStateTransitionAllowed := FInitialized AND
            (FState <> E_State.Uninitialized) AND (FState <> E_State.Reset) AND
            (FState <> E_State.Idle) AND (FState <> E_State.Completed);
ELSE
    IsStateTransitionAllowed := FALSE;
END_CASE;

IF ((NewState >= E_State.Preparing) AND (NewState < E_State.Completing)) AND
    ((FResult = E_Result.Error) OR (FAggregator.Result = E_Result.Error)) THEN
    IsStateTransitionAllowed := FALSE;
END_IF;
END_METHOD

{region 'Documentation'}
(*!
<summary>Reports Starting, configured Preparation/Test states, abort handling, legacy Aborted, or
Completing.</summary>
*)
{endregion}
{attribute 'monitoring' := 'call'}
PROPERTY PUBLIC IsTestCaseActive : BOOL //! Reports Starting, configured Preparation/Test states, abort handling, legacy Aborted, or Completing.
GET // PUBLIC
IsTestCaseActive := (FState = E_State.Starting) OR IsPreparationActive OR IsTestingActive
    OR (FState = E_State.Aborting) OR (FState = E_State.AbortingFromError) OR (FState = E_State.Aborted) OR (FState = E_State.Completing);
END_GET
END_PROPERTY

{region 'Documentation'}
(*!
<summary>Reports membership in the configured Test-state interval.</summary>
*)
{endregion}
{attribute 'monitoring' := 'call'}
PROPERTY PUBLIC IsTestingActive : BOOL //! Reports membership in the configured Test-state interval.
GET // PUBLIC
IsTestingActive := (FState >= E_State.Running) AND (FState < E_State.Running + FTestStateCount);
END_GET
END_PROPERTY

{region 'Documentation'}
(*!
<summary>Length-limited hierarchical name assigned by Initialize, including invalid diagnostic
names.</summary>
<description>
IsInitialized indicates successful initialization.
</description>
*)
{endregion}
{attribute 'monitoring' := 'variable'}
PROPERTY PUBLIC Name : STRING(GVL_Constants.NameLength) //! Length-limited hierarchical name assigned by Initialize, including invalid diagnostic names.
GET // PUBLIC
Name := FName;
END_GET
END_PROPERTY

{region 'Documentation'}
(*!
<summary>Advances immediately to the next configured Preparation state.</summary>
<description>
Only valid within the configured Preparation interval and without owner, aggregate or
Preparation Error. Advancing beyond the interval reports Error; use CompletePreparations to finish
the phase. The next state's timer starts with the transition.
</description>
*)
{endregion}
METHOD PROTECTED NextPreparationState
IF NOT IsPreparationActive THEN
    Error(Message := 'NextPreparationState called outside its lifecycle phase.');
    RETURN;
END_IF;
IF (FResult = E_Result.Error) OR (FAggregator.Result = E_Result.Error) THEN
    Error(Message := 'Test Case evaluation reported Error.');
    RETURN;
END_IF;

IF FState + 1 >= E_State.Preparing + FPreparationStateCount THEN
    Error(Message := 'NextPreparationState exceeds its configured state range.');
    RETURN;
END_IF;
IF FPreparationStatus.Error THEN
    Error(Message := 'Preparation reported Error.');
    RETURN;
END_IF;
ChangeState(NewState := FState + 1);
END_METHOD

{region 'Documentation'}
(*!
<summary>Advances immediately to the next configured Test state.</summary>
<description>
Only valid within the configured Test interval and without owner or aggregate Error. Advancing
beyond the interval reports Error; use CompleteTests to finish the phase. Later hooks in the same
call observe the new state.
</description>
*)
{endregion}
METHOD PROTECTED NextTestState
IF NOT IsTestingActive THEN
    Error(Message := 'NextTestState called outside its lifecycle phase.');
    RETURN;
END_IF;
IF (FResult = E_Result.Error) OR (FAggregator.Result = E_Result.Error) THEN
    Error(Message := 'Test Case evaluation reported Error.');
    RETURN;
END_IF;

IF FState + 1 >= E_State.Running + FTestStateCount THEN
    Error(Message := 'NextTestState exceeds its configured state range.');
    RETURN;
END_IF;
ChangeState(NewState := FState + 1);
END_METHOD

{region 'Documentation'}
(*!
<summary>Reports the configured maximum number of Preparation-state entries along one finite
lifecycle path.</summary>
<description>
Set the backing field explicitly in Configure. Before configuration it is
StateCountNotConfigured (-1). Branches use the longest path, including bounded repeated entries;
this is not a count of child instances. Keep it fixed through execution.

Zero means no Preparation phase. CheckInitialization bounds the value by E_State.Running -
E_State.Preparing.
</description>
*)
{endregion}
{attribute 'monitoring' := 'call'}
PROPERTY PUBLIC PreparationStateCount : INT //! Reports the configured maximum number of Preparation-state entries along one finite lifecycle path.
GET // PUBLIC
PreparationStateCount := FPreparationStateCount;
END_GET
END_PROPERTY

{region 'Documentation'}
(*!
<summary>Returns the stored combined Preparation observations without executing children.</summary>
*)
{endregion}
PROPERTY PUBLIC PreparationStatus : ST_PreparationStatus //! Returns the stored combined Preparation observations without executing children.
GET // PUBLIC
PreparationStatus := FPreparationStatus;
END_GET
END_PROPERTY

{region 'Documentation'}
(*!
<summary>Performs scenario cleanup during explicit or error-driven abort.</summary>
<description>
Called before Preparation and Test hooks on every initialized call except Completed. Enable is
TRUE only in an abort phase; disabled calls must not advance it.

Call CompleteAbort when cleanup is finished. The base owns the abort deadline, including
escalation from Abort to Error. This abstract hook has no base implementation.
</description>
*)
{endregion}
METHOD PROTECTED ABSTRACT ProcessAbort
VAR_INPUT
    Enable: BOOL; //! TRUE while this hook's lifecycle phase is active; FALSE must not advance that phase.
END_VAR
(* Example: process cleanup on enabled and disabled calls as required.
MyCleanup(Enable := Enable);
IF Enable AND MyCleanup.Completed THEN
    CompleteAbort();
END_IF;
*)
END_METHOD

{region 'Documentation'}
(*!
<summary>Executes owned Assertions with their current inputs and effective activation.</summary>
<description>
Called after ProcessTests on every initialized call except Completed. Enable is recomputed
from the current Test state, so CompleteTests earlier in the call disables enable-controlled
observation.

Keep disabled calls needed for pending resets and history; explicitly gated Evaluate inputs
remain the concrete scenario's responsibility. Result collection belongs to AggregateResults, not
this hook. This abstract hook has no base implementation.
</description>
*)
{endregion}
METHOD PROTECTED ABSTRACT ProcessAssertions
VAR_INPUT
    Enable: BOOL; //! TRUE while this hook's lifecycle phase is active; FALSE must not advance that phase.
END_VAR
(* Example: call each owned Assertion, including when Enable is FALSE.
MyAssertion(Enable := Enable,
    IN := ActualValue,
    Expected := ExpectedValue);
*)
END_METHOD

